(* PLC project HomeAutomation.ecp, WAGO e!COCKPIT e!COCKPIT *)
(* stored: creationDateTime 2023-02-09T18:04:59.3386506, modificationDateTime 2023-02-09T18:04:38.0443981 *)

{attribute 'to_string'}
TYPE Dimmer : (idle, soft_turn_on_restore, soft_turn_off, quick_turn_on, quick_turn_off, ramp_up_or_down, low_or_high_entering, low_or_high_leaving, low_or_high_released_by_user, blink);
END_TYPE

TYPE DIMMER_CURVE : (linear, logarithmic, cubic);
END_TYPE

TYPE MQTT_DISCOVERY_BASE : STRUCT
  name : JSONVAR;
  obj_id : JSONVAR;  (* object_id *)
  uniq_id : JSONVAR;  (* unique_id *)
  avty_t : JSONVAR;  (* availability_topic *)
  pl_avail : JSONVAR;  (* payload_available *)
  pl_not_avail : JSONVAR;  (* payload_not_available *)
  dev : MQTT_DISCOVERY_DEVICE;  (* device *)
  meta : JSONVAR;  (* extra metadata *)
END_STRUCT;
END_TYPE

TYPE MQTT_DISCOVERY_BINARY_SENSOR : STRUCT
  stat_t : JSONVAR;  (* state_topic *)
  pl_on : JSONVAR;  (* payload_on *)
  pl_off : JSONVAR;  (* payload_off *)
  dev_cla : JSONVAR;  (* device class *)
END_STRUCT;
END_TYPE

TYPE MQTT_DISCOVERY_COVER : STRUCT
  cmd_t : JSONVAR;  (* command_topic *)
  pl_open : JSONVAR;  (* payload open *)
  pl_cls : JSONVAR;  (* payload_close *)
  pl_stop : JSONVAR;  (* payload_stop *)
  stat_t : JSONVAR;  (* state topic *)
  stat_open : JSONVAR;  (* state open *)
  stat_clsd : JSONVAR;  (* state closed *)
  opt : JSONVAR;  (* optimistic *)
  dev_cla : JSONVAR;  (* device class *)
END_STRUCT;
END_TYPE

TYPE MQTT_DISCOVERY_DEVICE : STRUCT
  name : JSONVAR;
  cu : JSONVAR;  (* configuration_url *)
  ids : JSONVAR;  (* identifiers *)
  mf : JSONVAR;  (* manufacturer *)
  mdl : JSONVAR;  (* model *)
  sw : JSONVAR;  (* sw_version *)
  hw : JSONVAR;  (* hw_version *)
END_STRUCT;
END_TYPE

TYPE MQTT_DISCOVERY_LIGHT : STRUCT
  cmd_t : JSONVAR;  (* command_topic *)
  pl_on : JSONVAR;  (* payload_on *)
  pl_off : JSONVAR;  (* payload_off *)
  stat_t : JSONVAR;  (* state_topic *)
  opt : JSONVAR;  (* optimistic *)
END_STRUCT;
END_TYPE

TYPE MQTT_DISCOVERY_LIGHT_DIMMER : STRUCT
  bri_stat_t : JSONVAR;  (* brightness state topic *)
  bri_cmd_t : JSONVAR;  (* brightness command topic *)
  bri_scl : JSONVAR;  (* brightness scale *)
  on_cmd_type : JSONVAR;  (* on command type *)
  dmxChannel : JSONVAR;  (* DMX *)
  dmxWidth : JSONVAR;
  dmxUniverse : JSONVAR;
END_STRUCT;
END_TYPE

TYPE MQTT_DISCOVERY_LOCK : STRUCT
  cmd_t : JSONVAR;  (* command_topic *)
  pl_lock : JSONVAR;  (* payload lock *)
  pl_unlk : JSONVAR;  (* payload unlock *)
  stat_t : JSONVAR;  (* state_topic *)
  stat_locked : JSONVAR;  (* state locked *)
  stat_unlocked : JSONVAR;  (* state unlocked *)
  opt : JSONVAR;  (* optimistic *)
END_STRUCT;
END_TYPE

TYPE MQTT_DISCOVERY_SENSOR : STRUCT
  stat_t : JSONVAR;  (* state_topic *)
  exp_aft : JSONVAR;  (* expire after *)
END_STRUCT;
END_TYPE

TYPE MQTT_DISCOVERY_SIREN : STRUCT
  cmd_t : JSONVAR;  (* command_topic *)
  pl_on : JSONVAR;  (* payload_on *)
  pl_off : JSONVAR;  (* payload_off *)
  stat_t : JSONVAR;  (* state_topic *)
  stat_on : JSONVAR;  (* state on *)
  stat_off : JSONVAR;  (* state off *)
  opt : JSONVAR;  (* optimistic *)
END_STRUCT;
END_TYPE

TYPE MQTT_DISCOVERY_SWITCH : STRUCT
  cmd_t : JSONVAR;  (* command_topic *)
  pl_on : JSONVAR;  (* payload_on *)
  pl_off : JSONVAR;  (* payload_off *)
  stat_t : JSONVAR;  (* state_topic *)
  stat_on : JSONVAR;  (* state on *)
  stat_off : JSONVAR;  (* state off *)
  opt : JSONVAR;  (* optimistic *)
  dev_cla : JSONVAR;  (* device class *)
END_STRUCT;
END_TYPE

TYPE MQTT_MESSAGE : STRUCT
  Payload : STRING(1500);
  Topic : STRING(128);
  Qos : MQTT.QoS;
  MqttRetain : BOOL;
END_STRUCT;
END_TYPE

TYPE RS485_EASTRON_SDM_Devices : (SDM120, SDM220, SDM630);
END_TYPE

TYPE RS485_RtuQuery : STRUCT
  DeviceId : BYTE;
  FunctionCode : BYTE;
  ReadAddress : UINT;
  ReadQuantity : UINT;
  WriteAddress : UINT;
  WriteQuantity : UINT;
  WriteData : ARRAY[0..124] OF WORD;
END_STRUCT;
END_TYPE

TYPE VIRTUAL_MODES : (Input, Output);
END_TYPE

INTERFACE RS485Device
METHOD RequestBusTime : BOOL
END_METHOD
METHOD GetRtuQuery : RS485_RtuQuery
END_METHOD
METHOD ProcessDataArray
  VAR_INPUT
    Error : POINTER TO BOOL;
    Data : POINTER TO ARRAY[0..124] OF WORD;
  END_VAR
END_METHOD
END_INTERFACE

{attribute 'reflection'}
FUNCTION_BLOCK FB_BASE_MQTT_DISCOVERY_DEVICE
  VAR
    name : STRING;
    cu : STRING;  (* configuration_url *)
    cns : ARRAY[1..2] OF ARRAY[1..2] OF STRING;  (* connections *)
    ids : STRING;  (* identifiers *)
    mf : STRING;  (* manufacturer *)
    mdl : STRING;  (* model *)
    sw : STRING;  (* sw_version *)
    hw : STRING;  (* hw_version *)
    ip : STRING;
    mac : STRING;
    sAppName : STRING := 'Application';  (* must identic to the name in the device tree *)
    iecResult : RTS_IEC_RESULT;
    xInit : BOOL := TRUE;
    pApp : POINTER TO CmpApp.APPLICATION;
    stAppInfo : CmpApp.APPLICATION_INFO;
    pstAppInfo : POINTER TO CmpApp.APPLICATION_INFO := ADR(stAppInfo);
    {attribute 'instance-path'}
    {attribute 'noinit'}
    InstanceName : STRING;  (* object's full instance name *)
    Startup : BOOL := TRUE;
    InitMqttDone : BOOL;
    pMqttPublishQueue : POINTER TO FB_MqttPublishQueue;
    availabilityTopic : STRING;
    availabilityOnline : STRING;
    availabilityOffline : STRING;
    MqttDiscoveryPrefix : STRING;
    MqttDiscMsgBinSens : MQTT_DISCOVERY_BINARY_SENSOR;
    MqttDiscMsgCover : MQTT_DISCOVERY_COVER;
    MqttDiscMsgLightDim : MQTT_DISCOVERY_LIGHT_DIMMER;
    MqttDiscMsgLight : MQTT_DISCOVERY_LIGHT;
    MqttDiscMsgLock : MQTT_DISCOVERY_LOCK;
    MqttDiscMsgSensor : MQTT_DISCOVERY_SENSOR;
    MqttDiscMsgSiren : MQTT_DISCOVERY_SIREN;
    MqttDiscMsgSwitch : MQTT_DISCOVERY_SWITCH;
  END_VAR

            
          

{attribute 'reflection'}
METHOD CreateBinarySensorEntity
  VAR_INPUT
    Name : STRING;  (* default *)
    Id : STRING;
    Meta : STRING;
    StateTopic : STRING;  (* entity specific *)
    PayloadOn : STRING;
    PayloadOff : STRING;
    DeviceClass : STRING;
  END_VAR
  VAR
    EntityId : STRING(25) := 'binary_sensor';
    ComposeJSON : STRUCT_TO_JSON;
    MqttJSON : STRING(1500);
    MqttTopic : STRING(100);
  END_VAR
                  MqttTopic := CONCAT(CONCAT(CONCAT(CONCAT(THIS^.MqttDiscoveryPrefix, EntityId),'/'), Id),'/config' );


// 	Entity related: Basis
MqttDiscMsgBinSens.name.CharString :=  name; // friendly name
MqttDiscMsgBinSens.obj_id.CharString :=  Id; 
MqttDiscMsgBinSens.uniq_id.CharString :=  Id; 

// Entity related: Specific
MqttDiscMsgBinSens.stat_t.CharString := StateTopic;
MqttDiscMsgBinSens.pl_on.CharString := PayloadOn;
MqttDiscMsgBinSens.pl_off.CharString := PayloadOff;
MqttDiscMsgBinSens.dev_cla.CharString := DeviceClass;

// Availabilty related
MqttDiscMsgBinSens.avty_t.CharString :=  THIS^.availabilityTopic;
MqttDiscMsgBinSens.pl_avail.CharString :=   THIS^.availabilityOnline;
MqttDiscMsgBinSens.pl_not_avail.CharString :=  THIS^.availabilityOffline;

// Device related
MqttDiscMsgBinSens.dev.cu.CharString := THIS^.cu;
MqttDiscMsgBinSens.dev.name.CharString := THIS^.name;
MqttDiscMsgBinSens.dev.hw.CharString := THIS^.hw;
MqttDiscMsgBinSens.dev.ids.CharString := THIS^.ids;
MqttDiscMsgBinSens.dev.sw.CharString := THIS^.sw;
MqttDiscMsgBinSens.dev.mdl.CharString := THIS^.mdl;
MqttDiscMsgBinSens.dev.mf.CharString := THIS^.mf;
	
// Extra meta-data
IF NOT CommonTypesAndFunctions.StrEquals(str1:= ADR(meta), str2:= ADR('')) THEN
	MqttDiscMsgBinSens.meta.CharString := meta;
END_IF

ComposeJSON(
	JSONString:= ADR(MqttJSON), 
	JSONStringSize:= SIZEOF(MqttJSON),
	JSONVars:= ADR(MqttDiscMsgBinSens),
	NumberOfVars:= SIZEOF(MqttDiscMsgBinSens) / SIZEOF(JSONVAR),
	MaxLevel := 1,
);
ComposeJSON.Execute := TRUE;
ComposeJSON();

IF MqttJSON = '' THEN
	Mqttvariables.MQTT_logger.send(str:=CONCAT(CONCAT('ERROR ',Id), ' had empty MqttJSON'), instance := 'bla');
ELSIF NOT (MqttJSON = '') THEN
	pMqttPublishQueue^.AddMessage(
		Payload:= MqttJSON,
		Topic := MqttTopic,
		Qos := MQTT.QoS.ExactlyOnce,
		MqttRetain := TRUE,
	);
	Mqttvariables.MQTT_logger.send(str:=CONCAT(CONCAT('Added ',Id), ' as MQTT dicovery'), instance := 'bla');
END_IF

                
END_METHOD

METHOD CreateCoverEntity
  VAR_INPUT
    Name : STRING;  (* default *)
    Id : STRING;
    Meta : STRING;
    CommandTopic : STRING;  (* entity specific *)
    PayloadOpen : STRING;
    PayloadClose : STRING;
    PayloadStop : STRING;
    StateTopic : STRING;
    StateOpen : STRING;
    StateClosed : STRING;
    Deviceclass : STRING;
  END_VAR
  VAR
    EntityId : STRING(25) := 'cover';
    ComposeJSON : STRUCT_TO_JSON;
    MqttJSON : STRING(1500);
    MqttTopic : STRING(100);
  END_VAR
                  MqttTopic := CONCAT(CONCAT(CONCAT(CONCAT(THIS^.MqttDiscoveryPrefix, EntityId),'/'), Id),'/config' );

// 	Entity related: Basis
MqttDiscMsgCover.name.CharString :=  name; // friendly name
MqttDiscMsgCover.obj_id.CharString :=  Id; 
MqttDiscMsgCover.uniq_id.CharString :=  Id; 

// Entity related: Specific
MqttDiscMsgCover.cmd_t.CharString := CommandTopic;
MqttDiscMsgCover.pl_open.CharString := PayloadOpen;
MqttDiscMsgCover.pl_cls.CharString := PayloadClose;
MqttDiscMsgCover.pl_stop.CharString := PayloadStop;
MqttDiscMsgCover.stat_t.CharString := StateTopic;
MqttDiscMsgCover.stat_open.CharString := StateOpen;
MqttDiscMsgCover.stat_clsd.CharString := StateClosed;
MqttDiscMsgCover.opt.Boolean := FALSE;
MqttDiscMsgCover.dev_cla.CharString := Deviceclass;

// Availabilty related
MqttDiscMsgCover.avty_t.CharString :=  THIS^.availabilityTopic;
MqttDiscMsgCover.pl_avail.CharString :=   THIS^.availabilityOnline;
MqttDiscMsgCover.pl_not_avail.CharString :=  THIS^.availabilityOffline;

// Device related
MqttDiscMsgCover.dev.cu.CharString := THIS^.cu;
MqttDiscMsgCover.dev.name.CharString := THIS^.name;
MqttDiscMsgCover.dev.hw.CharString := THIS^.hw;
MqttDiscMsgCover.dev.ids.CharString := THIS^.ids;
MqttDiscMsgCover.dev.sw.CharString := THIS^.sw;
MqttDiscMsgCover.dev.mdl.CharString := THIS^.mdl;
MqttDiscMsgCover.dev.mf.CharString := THIS^.mf;
	
// Extra meta-data
IF NOT CommonTypesAndFunctions.StrEquals(str1:= ADR(meta), str2:= ADR('')) THEN
	MqttDiscMsgCover.meta.CharString := meta;
END_IF

ComposeJSON(
	JSONString:= ADR(MqttJSON), 
	JSONStringSize:= SIZEOF(MqttJSON),
	JSONVars:= ADR(MqttDiscMsgCover),
	NumberOfVars:= SIZEOF(MqttDiscMsgCover) / SIZEOF(JSONVAR),
	MaxLevel := 1,
);
ComposeJSON.Execute := TRUE;
ComposeJSON();

IF MqttJSON = '' THEN
	Mqttvariables.MQTT_logger.send(str:=CONCAT(CONCAT('ERROR ',Id), ' had empty MqttJSON'), instance := 'bla');
ELSIF NOT (MqttJSON = '') THEN
	pMqttPublishQueue^.AddMessage(
		Payload:= MqttJSON,
		Topic := MqttTopic,
		Qos := MQTT.QoS.ExactlyOnce,
		MqttRetain := TRUE,
	);
	Mqttvariables.MQTT_logger.send(str:=CONCAT(CONCAT('Added ',Id), ' as MQTT dicovery'), instance := 'bla');
END_IF

                
END_METHOD

METHOD initBaseDevice
  VAR_INPUT
    Name : STRING;
    ConfigurationUrl : STRING;
    Identifiers : STRING;
    Manufacturer : STRING;
    Model : STRING;
    SoftwareVersion : STRING;
    HardwareVersion : STRING;
    IpAddress : STRING := '';
    MacAddress : STRING := '';
    availabilityTopic : STRING;
    availabilityOnline : STRING;
    availabilityOffline : STRING;
    MqttDiscoveryPrefix : STRING;
    pMqttPublishQueue : POINTER TO FB_MqttPublishQueue;
  END_VAR
                  THIS^.availabilityTopic := availabilityTopic;
THIS^.availabilityOnline := availabilityOnline;
THIS^.availabilityOffline := availabilityOffline;
THIS^.pMqttPublishQueue := pMqttPublishQueue;
THIS^.MqttDiscoveryPrefix := MqttDiscoveryPrefix;

THIS^.name := Name;
THIS^.cu:= ConfigurationUrl;
THIS^.ids:= Identifiers;
THIS^.mf:= Manufacturer;
THIS^.mdl:= Model;
THIS^.hw:= HardwareVersion;
THIS^.ip := IpAddress;
THIS^.mac := MacAddress;




                
END_METHOD

METHOD CreateLightEntity
  VAR_INPUT
    Name : STRING;  (* default *)
    Id : STRING;
    Meta : STRING;
    CommandTopic : STRING;  (* entity specific *)
    PayloadOn : STRING;
    PayloadOff : STRING;
    StateTopic : STRING;
  END_VAR
  VAR
    EntityId : STRING(25) := 'light';
    ComposeJSON : STRUCT_TO_JSON;
    MqttJSON : STRING(1500);
    MqttTopic : STRING(100);
  END_VAR
                  MqttTopic := CONCAT(CONCAT(CONCAT(CONCAT(THIS^.MqttDiscoveryPrefix, EntityId),'/'), Id),'/config' );

// 	Entity related: Basis
MqttDiscMsgLight.name.CharString :=  name; // friendly name
MqttDiscMsgLight.obj_id.CharString :=  Id; 
MqttDiscMsgLight.uniq_id.CharString :=  Id; 

// Entity related: Specific
MqttDiscMsgLight.cmd_t.CharString := CommandTopic;
MqttDiscMsgLight.pl_on.CharString := PayloadOn;
MqttDiscMsgLight.pl_off.CharString := PayloadOff;
MqttDiscMsgLight.stat_t.CharString := StateTopic;
MqttDiscMsgLight.opt.Boolean := FALSE;

// Availabilty related
MqttDiscMsgLight.avty_t.CharString :=  THIS^.availabilityTopic;
MqttDiscMsgLight.pl_avail.CharString :=   THIS^.availabilityOnline;
MqttDiscMsgLight.pl_not_avail.CharString :=  THIS^.availabilityOffline;

// Device related
MqttDiscMsgLight.dev.cu.CharString := THIS^.cu;
MqttDiscMsgLight.dev.name.CharString := THIS^.name;
MqttDiscMsgLight.dev.hw.CharString := THIS^.hw;
MqttDiscMsgLight.dev.ids.CharString := THIS^.ids;
MqttDiscMsgLight.dev.sw.CharString := THIS^.sw;
MqttDiscMsgLight.dev.mdl.CharString := THIS^.mdl;
MqttDiscMsgLight.dev.mf.CharString := THIS^.mf;
	
// Extra meta-data
IF NOT CommonTypesAndFunctions.StrEquals(str1:= ADR(meta), str2:= ADR('')) THEN
	MqttDiscMsgLight.meta.CharString := meta;
END_IF

ComposeJSON(
	JSONString:= ADR(MqttJSON), 
	JSONStringSize:= SIZEOF(MqttJSON),
	JSONVars:= ADR(MqttDiscMsgLight),
	NumberOfVars:= SIZEOF(MqttDiscMsgLight) / SIZEOF(JSONVAR),
	MaxLevel := 1,
);
ComposeJSON.Execute := TRUE;
ComposeJSON();

IF MqttJSON = '' THEN
	Mqttvariables.MQTT_logger.send(str:=CONCAT(CONCAT('ERROR ',Id), ' had empty MqttJSON'), instance := 'bla');
ELSIF NOT (MqttJSON = '') THEN
	pMqttPublishQueue^.AddMessage(
		Payload:= MqttJSON,
		Topic := MqttTopic,
		Qos := MQTT.QoS.ExactlyOnce,
		MqttRetain := TRUE,
	);
	Mqttvariables.MQTT_logger.send(str:=CONCAT(CONCAT('Added ',Id), ' as MQTT dicovery'), instance := 'bla');
END_IF

                
END_METHOD

METHOD CreateLockEntity
  VAR_INPUT
    Name : STRING;  (* default *)
    Id : STRING;
    Meta : STRING;
    CommandTopic : STRING;  (* entity specific *)
    PayloadLock : STRING;
    PayloadUnlock : STRING;
    StateTopic : STRING;
    StateLocked : STRING;
    StateUnlocked : STRING;
  END_VAR
  VAR
    EntityId : STRING(25) := 'lock';
    ComposeJSON : STRUCT_TO_JSON;
    MqttJSON : STRING(1500);
    MqttTopic : STRING(100);
  END_VAR
                  MqttTopic := CONCAT(CONCAT(CONCAT(CONCAT(THIS^.MqttDiscoveryPrefix, EntityId),'/'), Id),'/config' );

// 	Entity related: Basis
MqttDiscMsgLock.name.CharString :=  name; // friendly name
MqttDiscMsgLock.obj_id.CharString :=  Id; 
MqttDiscMsgLock.uniq_id.CharString :=  Id; 

// Entity related: Specific
MqttDiscMsgLock.cmd_t.CharString := CommandTopic;
MqttDiscMsgLock.pl_lock.CharString := PayloadLock;
MqttDiscMsgLock.pl_unlk.CharString := PayloadUnlock;
MqttDiscMsgLock.stat_t.CharString := StateTopic;
MqttDiscMsgLock.stat_locked.CharString := StateLocked;
MqttDiscMsgLock.stat_unlocked.CharString := StateUnlocked;
MqttDiscMsgLock.opt.Boolean := FALSE;

// Availabilty related
MqttDiscMsgLock.avty_t.CharString :=  THIS^.availabilityTopic;
MqttDiscMsgLock.pl_avail.CharString :=   THIS^.availabilityOnline;
MqttDiscMsgLock.pl_not_avail.CharString :=  THIS^.availabilityOffline;

// Device related
MqttDiscMsgLock.dev.cu.CharString := THIS^.cu;
MqttDiscMsgLock.dev.name.CharString := THIS^.name;
MqttDiscMsgLock.dev.hw.CharString := THIS^.hw;
MqttDiscMsgLock.dev.ids.CharString := THIS^.ids;
MqttDiscMsgLock.dev.sw.CharString := THIS^.sw;
MqttDiscMsgLock.dev.mdl.CharString := THIS^.mdl;
MqttDiscMsgLock.dev.mf.CharString := THIS^.mf;
	
// Extra meta-data
IF NOT CommonTypesAndFunctions.StrEquals(str1:= ADR(meta), str2:= ADR('')) THEN
	MqttDiscMsgLock.meta.CharString := meta;
END_IF

ComposeJSON(
	JSONString:= ADR(MqttJSON), 
	JSONStringSize:= SIZEOF(MqttJSON),
	JSONVars:= ADR(MqttDiscMsgLock),
	NumberOfVars:= SIZEOF(MqttDiscMsgLock) / SIZEOF(JSONVAR),
	MaxLevel := 1,
);
ComposeJSON.Execute := TRUE;
ComposeJSON();

IF MqttJSON = '' THEN
	Mqttvariables.MQTT_logger.send(str:=CONCAT(CONCAT('ERROR ',Id), ' had empty MqttJSON'), instance := 'bla');
ELSIF NOT (MqttJSON = '') THEN
	pMqttPublishQueue^.AddMessage(
		Payload:= MqttJSON,
		Topic := MqttTopic,
		Qos := MQTT.QoS.ExactlyOnce,
		MqttRetain := TRUE,
	);
	Mqttvariables.MQTT_logger.send(str:=CONCAT(CONCAT('Added ',Id), ' as MQTT dicovery'), instance := 'bla');
END_IF

                
END_METHOD

METHOD CreateSirenEntity
  VAR_INPUT
    Name : STRING;  (* default *)
    Id : STRING;
    Meta : STRING;
    CommandTopic : STRING;  (* entity specific *)
    PayloadOn : STRING;
    PayloadOff : STRING;
    StateTopic : STRING;
    StateOnPayload : STRING;
    StateOffPayload : STRING;
  END_VAR
  VAR
    EntityId : STRING(25) := 'siren';
    ComposeJSON : STRUCT_TO_JSON;
    MqttJSON : STRING(1500);
    MqttTopic : STRING(100);
  END_VAR
                  MqttTopic := CONCAT(CONCAT(CONCAT(CONCAT(THIS^.MqttDiscoveryPrefix, EntityId),'/'), Id),'/config' );

// 	Entity related: Basis
MqttDiscMsgSiren.name.CharString :=  name; // friendly name
MqttDiscMsgSiren.obj_id.CharString :=  Id; 
MqttDiscMsgSiren.uniq_id.CharString :=  Id; 

// Entity related: Specific
MqttDiscMsgSiren.cmd_t.CharString := CommandTopic;
MqttDiscMsgSiren.pl_on.CharString := PayloadOn;
MqttDiscMsgSiren.pl_off.CharString := PayloadOff;
MqttDiscMsgSiren.stat_t.CharString := StateTopic;
MqttDiscMsgSiren.stat_on.CharString := StateOnPayload;
MqttDiscMsgSiren.stat_off.CharString := StateOffPayload;
MqttDiscMsgSiren.opt.Boolean := FALSE;

// Availabilty related
MqttDiscMsgSiren.avty_t.CharString :=  THIS^.availabilityTopic;
MqttDiscMsgSiren.pl_avail.CharString :=   THIS^.availabilityOnline;
MqttDiscMsgSiren.pl_not_avail.CharString :=  THIS^.availabilityOffline;

// Device related
MqttDiscMsgSiren.dev.cu.CharString := THIS^.cu;
MqttDiscMsgSiren.dev.name.CharString := THIS^.name;
MqttDiscMsgSiren.dev.hw.CharString := THIS^.hw;
MqttDiscMsgSiren.dev.ids.CharString := THIS^.ids;
MqttDiscMsgSiren.dev.sw.CharString := THIS^.sw;
MqttDiscMsgSiren.dev.mdl.CharString := THIS^.mdl;
MqttDiscMsgSiren.dev.mf.CharString := THIS^.mf;
	
// Extra meta-data
IF NOT CommonTypesAndFunctions.StrEquals(str1:= ADR(meta), str2:= ADR('')) THEN
	MqttDiscMsgSiren.meta.CharString := meta;
END_IF

ComposeJSON(
	JSONString:= ADR(MqttJSON), 
	JSONStringSize:= SIZEOF(MqttJSON),
	JSONVars:= ADR(MqttDiscMsgSiren),
	NumberOfVars:= SIZEOF(MqttDiscMsgSiren) / SIZEOF(JSONVAR),
	MaxLevel := 1,
);
ComposeJSON.Execute := TRUE;
ComposeJSON();

IF MqttJSON = '' THEN
	Mqttvariables.MQTT_logger.send(str:=CONCAT(CONCAT('ERROR ',Id), ' had empty MqttJSON'), instance := 'bla');
ELSIF NOT (MqttJSON = '') THEN
	pMqttPublishQueue^.AddMessage(
		Payload:= MqttJSON,
		Topic := MqttTopic,
		Qos := MQTT.QoS.ExactlyOnce,
		MqttRetain := TRUE,
	);
	Mqttvariables.MQTT_logger.send(str:=CONCAT(CONCAT('Added ',Id), ' as MQTT dicovery'), instance := 'bla');
END_IF

                
END_METHOD

METHOD CreateSensorEntity
  VAR_INPUT
    Name : STRING;  (* default *)
    Id : STRING;
    Meta : STRING;
    StateTopic : STRING;  (* entity specific *)
    ExpiryAfter : INT := 0;
  END_VAR
  VAR
    EntityId : STRING(25) := 'sensor';
    ComposeJSON : STRUCT_TO_JSON;
    MqttJSON : STRING(1500);
    MqttTopic : STRING(100);
  END_VAR
                  MqttTopic := CONCAT(CONCAT(CONCAT(CONCAT(THIS^.MqttDiscoveryPrefix, EntityId),'/'), Id),'/config' );

// 	Entity related: Basis
MqttDiscMsgSensor.name.CharString :=  name; // friendly name
MqttDiscMsgSensor.obj_id.CharString :=  Id; 
MqttDiscMsgSensor.uniq_id.CharString :=  Id; 

// Entity related: Specific
//MqttDiscoverySensorMessage.ic.CharString := Icon;
MqttDiscMsgSensor.stat_t.CharString := StateTopic;
MqttDiscMsgSensor.exp_aft.Integer := ExpiryAfter;

// Availabilty related
MqttDiscMsgSensor.avty_t.CharString :=  THIS^.availabilityTopic;
MqttDiscMsgSensor.pl_avail.CharString :=   THIS^.availabilityOnline;
MqttDiscMsgSensor.pl_not_avail.CharString :=  THIS^.availabilityOffline;

// Device related
MqttDiscMsgSensor.dev.cu.CharString := THIS^.cu;
MqttDiscMsgSensor.dev.name.CharString := THIS^.name;
MqttDiscMsgSensor.dev.hw.CharString := THIS^.hw;
MqttDiscMsgSensor.dev.ids.CharString := THIS^.ids;
MqttDiscMsgSensor.dev.sw.CharString := THIS^.sw;
MqttDiscMsgSensor.dev.mdl.CharString := THIS^.mdl;
MqttDiscMsgSensor.dev.mf.CharString := THIS^.mf;
	
// Extra meta-data
IF NOT CommonTypesAndFunctions.StrEquals(str1:= ADR(meta), str2:= ADR('')) THEN
	MqttDiscMsgSensor.meta.CharString := meta;
END_IF

ComposeJSON(
	JSONString:= ADR(MqttJSON), 
	JSONStringSize:= SIZEOF(MqttJSON),
	JSONVars:= ADR(MqttDiscMsgSensor),
	NumberOfVars:= SIZEOF(MqttDiscMsgSensor) / SIZEOF(JSONVAR),
	MaxLevel := 1,
);
ComposeJSON.Execute := TRUE;
ComposeJSON();

IF MqttJSON = '' THEN
	Mqttvariables.MQTT_logger.send(str:=CONCAT(CONCAT('ERROR ',Id), ' had empty MqttJSON'), instance := 'bla');
ELSIF NOT (MqttJSON = '') THEN
	pMqttPublishQueue^.AddMessage(
		Payload:= MqttJSON,
		Topic := MqttTopic,
		Qos := MQTT.QoS.ExactlyOnce,
		MqttRetain := TRUE,
	);
	Mqttvariables.MQTT_logger.send(str:=CONCAT(CONCAT('Added ',Id), ' as MQTT dicovery'), instance := 'bla');
END_IF

                
END_METHOD

METHOD CreateLightDimmerEntity
  VAR_INPUT
    Name : STRING;  (* default *)
    Id : STRING;
    Meta : STRING;
    CommandTopic : STRING;  (* entity specific *)
    PayloadOn : STRING;
    PayloadOff : STRING;
    StateTopic : STRING;
    BrightnessCommandTopic : STRING;
    BrightnessStateTopic : STRING;
    BrightnessScale : INT;
    DmxChannel : INT := 0;  (* dmx specific *)
    DmxWidth : INT := 0;
    DmxUniverse : INT := 0;
  END_VAR
  VAR
    EntityId : STRING(25) := 'light';
    ComposeJSON : STRUCT_TO_JSON;
    MqttJSON : STRING(1500);
    MqttTopic : STRING(100);
  END_VAR
                  MqttTopic := CONCAT(CONCAT(CONCAT(CONCAT(THIS^.MqttDiscoveryPrefix, EntityId),'/'), Id),'/config' );

// 	Entity related: Basis
MqttDiscMsgLightDim.name.CharString :=  name; // friendly name
MqttDiscMsgLightDim.obj_id.CharString :=  Id; 
MqttDiscMsgLightDim.uniq_id.CharString :=  Id; 

// Entity related: Specific
MqttDiscMsgLightDim.cmd_t.CharString := CommandTopic;
MqttDiscMsgLightDim.pl_on.CharString := PayloadOn;
MqttDiscMsgLightDim.pl_off.CharString := PayloadOff;
MqttDiscMsgLightDim.stat_t.CharString := StateTopic;
MqttDiscMsgLightDim.opt.Boolean := FALSE;

MqttDiscMsgLightDim.bri_cmd_t.CharString := BrightnessCommandTopic;
MqttDiscMsgLightDim.bri_stat_t.CharString := BrightnessStateTopic;
MqttDiscMsgLightDim.bri_scl.Integer := BrightnessScale;
MqttDiscMsgLightDim.on_cmd_type.CharString := 'last';

MqttDiscMsgLightDim.dmxChannel.Integer := DmxChannel;
MqttDiscMsgLightDim.dmxWidth.Integer := DmxWidth;
MqttDiscMsgLightDim.dmxUniverse.Integer := DmxUniverse;

// Availabilty related
MqttDiscMsgLightDim.avty_t.CharString :=  THIS^.availabilityTopic;
MqttDiscMsgLightDim.pl_avail.CharString :=   THIS^.availabilityOnline;
MqttDiscMsgLightDim.pl_not_avail.CharString :=  THIS^.availabilityOffline;

// Device related
MqttDiscMsgLightDim.dev.cu.CharString := THIS^.cu;
MqttDiscMsgLightDim.dev.name.CharString := THIS^.name;
MqttDiscMsgLightDim.dev.hw.CharString := THIS^.hw;
MqttDiscMsgLightDim.dev.ids.CharString := THIS^.ids;
MqttDiscMsgLightDim.dev.sw.CharString := THIS^.sw;
MqttDiscMsgLightDim.dev.mdl.CharString := THIS^.mdl;
MqttDiscMsgLightDim.dev.mf.CharString := THIS^.mf;
	
// Extra meta-data
IF NOT CommonTypesAndFunctions.StrEquals(str1:= ADR(meta), str2:= ADR('')) THEN
	MqttDiscMsgLightDim.meta.CharString := meta;
END_IF

ComposeJSON(
	JSONString:= ADR(MqttJSON), 
	JSONStringSize:= SIZEOF(MqttJSON),
	JSONVars:= ADR(MqttDiscMsgLightDim),
	NumberOfVars:= SIZEOF(MqttDiscMsgLightDim) / SIZEOF(JSONVAR),
	MaxLevel := 1,
);
ComposeJSON.Execute := TRUE;
ComposeJSON();

IF MqttJSON = '' THEN
	Mqttvariables.MQTT_logger.send(str:=CONCAT(CONCAT('ERROR ',Id), ' had empty MqttJSON'), instance := 'bla');
ELSIF NOT (MqttJSON = '') THEN
	pMqttPublishQueue^.AddMessage(
		Payload:= MqttJSON,
		Topic := MqttTopic,
		Qos := MQTT.QoS.ExactlyOnce,
		MqttRetain := TRUE,
	);
	Mqttvariables.MQTT_logger.send(str:=CONCAT(CONCAT('Added ',Id), ' as MQTT dicovery'), instance := 'bla');
END_IF

                
END_METHOD

METHOD CreateSwitchEntity
  VAR_INPUT
    Name : STRING;  (* default *)
    Id : STRING;
    Meta : STRING;
    CommandTopic : STRING;  (* entity specific *)
    PayloadOn : STRING;
    PayloadOff : STRING;
    StateTopic : STRING;
    StateOnPayload : STRING;
    StateOffPayload : STRING;
    DeviceClass : STRING;
  END_VAR
  VAR
    EntityId : STRING(25) := 'switch';
    ComposeJSON : STRUCT_TO_JSON;
    MqttJSON : STRING(1500);
    MqttTopic : STRING(100);
  END_VAR
                  MqttTopic := CONCAT(CONCAT(CONCAT(CONCAT(THIS^.MqttDiscoveryPrefix, EntityId),'/'), Id),'/config' );

// 	Entity related: Basis
MqttDiscMsgSwitch.name.CharString :=  name; // friendly name
MqttDiscMsgSwitch.obj_id.CharString :=  Id; 
MqttDiscMsgSwitch.uniq_id.CharString :=  Id; 

// Entity related: Specific
MqttDiscMsgSwitch.cmd_t.CharString := CommandTopic;
MqttDiscMsgSwitch.pl_on.CharString := PayloadOn;
MqttDiscMsgSwitch.pl_off.CharString := PayloadOff;
MqttDiscMsgSwitch.stat_t.CharString := StateTopic;
MqttDiscMsgSwitch.stat_on.CharString := StateOnPayload;
MqttDiscMsgSwitch.stat_off.CharString := StateOffPayload;
MqttDiscMsgSwitch.opt.Boolean := FALSE;
MqttDiscMsgSwitch.dev_cla.CharString := DeviceClass;

// Availabilty related
MqttDiscMsgSwitch.avty_t.CharString :=  THIS^.availabilityTopic;
MqttDiscMsgSwitch.pl_avail.CharString :=   THIS^.availabilityOnline;
MqttDiscMsgSwitch.pl_not_avail.CharString :=  THIS^.availabilityOffline;

// Device related
MqttDiscMsgSwitch.dev.cu.CharString := THIS^.cu;
MqttDiscMsgSwitch.dev.name.CharString := THIS^.name;
MqttDiscMsgSwitch.dev.hw.CharString := THIS^.hw;
MqttDiscMsgSwitch.dev.ids.CharString := THIS^.ids;
MqttDiscMsgSwitch.dev.sw.CharString := THIS^.sw;
MqttDiscMsgSwitch.dev.mdl.CharString := THIS^.mdl;
MqttDiscMsgSwitch.dev.mf.CharString := THIS^.mf;
	
// Extra meta-data
IF NOT CommonTypesAndFunctions.StrEquals(str1:= ADR(meta), str2:= ADR('')) THEN
	MqttDiscMsgSwitch.meta.CharString := meta;
END_IF

ComposeJSON(
	JSONString:= ADR(MqttJSON), 
	JSONStringSize:= SIZEOF(MqttJSON),
	JSONVars:= ADR(MqttDiscMsgSwitch),
	NumberOfVars:= SIZEOF(MqttDiscMsgSwitch) / SIZEOF(JSONVAR),
	MaxLevel := 1,
);
ComposeJSON.Execute := TRUE;
ComposeJSON();

IF MqttJSON = '' THEN
	Mqttvariables.MQTT_logger.send(str:=CONCAT(CONCAT('ERROR ',Id), ' had empty MqttJSON'), instance := 'bla');
ELSIF NOT (MqttJSON = '') THEN
	pMqttPublishQueue^.AddMessage(
		Payload:= MqttJSON,
		Topic := MqttTopic,
		Qos := MQTT.QoS.ExactlyOnce,
		MqttRetain := TRUE,
	);
	Mqttvariables.MQTT_logger.send(str:=CONCAT(CONCAT('Added ',Id), ' as MQTT dicovery'), instance := 'bla');
END_IF

                
END_METHOD
END_FUNCTION_BLOCK

{attribute 'reflection'}
FUNCTION_BLOCK FB_INPUT_BINARYSENSOR_MQTT EXTENDS FB_MQTT_BASE
  VAR_INPUT
    BS : BOOL;
  END_VAR
  VAR_OUTPUT
    Q : BOOL;  (* Follows the input but debounced *)
    EVENT : BOOL;  (* Event outputs only high for on clock cycle *)
    EVENT_R : BOOL;
    EVENT_F : BOOL;
  END_VAR
  VAR
    {attribute 'instance-path'}
    {attribute 'noinit'}
    InstancePath : STRING;  (* object's full instance name *)
    Startup : BOOL := TRUE;
    FB_DEBOUNCE : OSCAT_BUILDING.DEBOUNCE;  (* to debounce the physical input *)
    FB_R_TRIG : Standard.R_TRIG;  (* to detect a rising edge on the debounced signal *)
    FB_F_TRIG : Standard.F_TRIG;  (* to detect a falling edge on the debounced signal *)
    T_TurnOffDelay : TIME := TIME#0ms;
    FB_TurnOffDelayTimer : TOF;
    MqttDiscoveryMessage : MQTT_DISCOVERY_BINARY_SENSOR;
  END_VAR

            FB_DEBOUNCE(IN := BS,	
	TD := T#50MS, (* 2x cyle + 10ms *)
	PM := FALSE
	);
	
FB_TurnOffDelayTimer(IN:=FB_DEBOUNCE.Q,
	PT := T_TurnOffDelay,
	Q=>Q
	);

FB_R_TRIG(CLK := FB_TurnOffDelayTimer.Q);
FB_F_TRIG(CLK := FB_TurnOffDelayTimer.Q);

EVENT := FB_R_TRIG.Q OR FB_F_TRIG.Q;
EVENT_R := FB_R_TRIG.Q;
EVENT_F := FB_F_TRIG.Q;

IF (FB_R_TRIG.Q OR (Startup AND FB_DEBOUNCE.Q)) AND InitMqttDone THEN
	pMqttPublishQueue^.AddMessage(
		Payload := 'ON',
		Topic := CONCAT(MqttPublishTopicPrefix^, MqttPublishTopicSuffix),
		Qos := MQTT.QoS.ExactlyOnce,
		MqttRetain := TRUE
	);
	Startup:=FALSE;	
END_IF

IF (FB_F_TRIG.Q OR (Startup AND NOT(FB_DEBOUNCE.Q))) AND InitMqttDone THEN
	pMqttPublishQueue^.AddMessage(
		Payload := 'OFF',
		Topic := CONCAT(MqttPublishTopicPrefix^, MqttPublishTopicSuffix),
		Qos := MQTT.QoS.ExactlyOnce,
		MqttRetain := TRUE
	);
	Startup:=FALSE;	
END_IF
          

METHOD InitMqtt
  VAR_INPUT
    MQTTPublishPrefix : POINTER TO STRING;
    pMqttPublishQueue : POINTER TO FB_MqttPublishQueue;
  END_VAR
                  SUPER^._InstancePath := THIS^.InstancePath; // Due to reflection its location is important

(*pass trough*)
THIS^.pMqttPublishQueue := pMqttPublishQueue;
THIS^.MqttPublishTopicPrefix:=MQTTPublishPrefix;
SUPER^.InitBaseMqtt();

                
END_METHOD

METHOD InitMqttDiscovery
  VAR_INPUT
    Device : POINTER TO FB_PLC_MQTT_DISCOVERY_DEVICE;
    Name : STRING(255);
    DeviceClass : STRING(100) := 'smoke';
    overruleId : STRING(255) := '';
    meta : STRING(255) := '';
  END_VAR
  VAR
    id : STRING(255);
  END_VAR
                  IF InitMqttDone AND NOT initMqttDiscoveryDone THEN
	
	IF CommonTypesAndFunctions.StrEquals(str1:= ADR(overruleId), str2:= ADR('')) THEN
		id := CONCAT(CONCAT(THIS^.DeviceName,'_'), THIS^.InstanceNamePt^); // 'FB_DI_PB_003'
	ELSE
		id := overruleId; // 'MY_PH_GND_HALL_01'
	END_IF
	
	Device^.CreateBinarySensorEntity(
		Id := id,
		Name := name,
		Meta := meta,
		StateTopic := THIS^.MQTTPublishTopic,
		PayloadOn := 'ON',
		PayloadOff := 'OFF',
		DeviceClass := DeviceClass);
		
	initMqttDiscoveryDone := TRUE;
END_IF		
                
END_METHOD

METHOD ConfigureFunctionBlock
  VAR_INPUT
    T_TurnOffDelay : TIME;
  END_VAR
                  THIS^.T_TurnOffDelay:=T_TurnOffDelay;
                
END_METHOD
END_FUNCTION_BLOCK

{attribute 'reflection'}
FUNCTION_BLOCK FB_INPUT_PUSHBUTTON_DIMMER_MQTT
  VAR_INPUT
    PB : BOOL;
    SET : BOOL;
    VAL : BYTE;
    RST : BOOL;
  END_VAR
  VAR_OUTPUT
    DIM : BYTE;
    DBL : BOOL;
    Q : BOOL;
    SINGLE : BOOL;
    DOUBLE : BOOL;
    LONG : BOOL;
    P_LONG : BOOL;
  END_VAR
  VAR
    {attribute 'instance-path'}
    {attribute 'noinit'}
    InstanceName : STRING;  (* object's full instance name *)
    InitMqttDone : BOOL;
    MqttPublishTopicPrefix : POINTER TO STRING;
    MqttPublishTopicSuffix : STRING(50);
    pMqttPublishQueue : POINTER TO FB_MqttPublishQueue;
    FB_DIMMER : OSCAT_BUILDING.DIMM_I;
    OutputDimmer : BOOL;
    Qos_Dimm : MQTT.QoS;
    Delta_Dimm : INT;
    FB_DETECTPUSH : OSCAT_BUILDING.CLICK_MODE;
    P_LONG_R_TRIG : Standard.R_TRIG;
    P_LONG_F_TRIG : Standard.F_TRIG;
    PreviousDim : BYTE;  (* Vars to detect statechanges on outputs *)
    PreviousQ : BOOL;
    PreviousDBL : BOOL;
    T_Debounce : TIME := TIME#10ms;  (* Default values for dimmer, can be overwritten by method call *)
    T_Reconfig : TIME := TIME#10s0ms;
    T_On_Max : TIME := TIME#0ms;
    T_Dimm_Start : TIME := TIME#400ms;
    T_Dimm : TIME := TIME#3s0ms;
    Min_On : BYTE := 50;
    Max_On : BYTE := 255;
    Soft_Dimm : BOOL := TRUE;
    Dbl_Toggle : BOOL := FALSE;
    Rst_Out : BOOL := FALSE;
    T_Long : TIME := TIME#400ms;  (* Default value for click mode, can be overwritten by method call *)
  END_VAR

            FB_DIMMER(
	IN:= PB,
	SET:= SET,
	VAL:= VAL,
	RST:= RST,
	OUT:= DIM,
	T_DEBOUNCE:= T_Debounce,
	T_RECONFIG:= T_Reconfig,
	T_ON_MAX:= T_On_Max,
	T_DIMM_START:= T_Dimm_Start,
	T_DIMM:= T_Dimm,
	MIN_ON:= Min_On,
	MAX_ON:= Max_On,
	SOFT_DIMM:= Soft_Dimm,
	DBL_TOGGLE:= Dbl_Toggle,
	RST_OUT:= Rst_Out,
	Q=> Q,
	DBL=> DBL);
	
FB_DETECTPUSH(
	IN:= PB, 	
	SINGLE=> SINGLE, 
	DOUBLE=> DOUBLE, 
	TP_LONG=> LONG, 
	T_LONG:= T_long);
	
P_LONG_R_TRIG(CLK:=FB_DETECTPUSH.LONG);
P_LONG_F_TRIG(CLK:=FB_DETECTPUSH.LONG);
	
IF (ABS(BYTE_TO_INT(PreviousDim) - BYTE_TO_INT(DIM)) >= Delta_Dimm OR PB = FALSE) AND DIM <> PreviousDim AND OutputDimmer AND InitMqttDone  THEN
	PreviousDim:=DIM;
	pMqttPublishQueue^.AddMessage(		
		Payload := BYTE_TO_STRING(DIM),
		Topic := CONCAT(CONCAT(MqttPublishTopicPrefix^, MqttPublishTopicSuffix), '/DIM'),
		Qos := MQTT.QoS.ExactlyOnce,
		MqttRetain := FALSE
	);
END_IF

IF FB_DIMMER.Q <> PreviousQ AND InitMqttDone THEN
	PreviousQ:=FB_DIMMER.Q;
	pMqttPublishQueue^.AddMessage(
		Payload := BOOL_TO_STRING(FB_DIMMER.Q),
		Topic := CONCAT(CONCAT(MqttPublishTopicPrefix^, MqttPublishTopicSuffix), '/Q'),
		Qos := Qos_Dimm,
		MqttRetain := TRUE
	);
END_IF

IF FB_DIMMER.DBL <> PreviousDBL AND InitMqttDone THEN
	PreviousDBL:=FB_DIMMER.DBL;
	pMqttPublishQueue^.AddMessage(
		Payload := BOOL_TO_STRING(FB_DIMMER.DBL),
		Topic := CONCAT(CONCAT(MqttPublishTopicPrefix^, MqttPublishTopicSuffix), '/DBL'),
		Qos := MQTT.QoS.ExactlyOnce,
		MqttRetain := TRUE
	);
END_IF

IF FB_DETECTPUSH.SINGLE AND InitMqttDone THEN
	pMqttPublishQueue^.AddMessage(
		Payload := 'SINGLE',
		Topic := CONCAT(MqttPublishTopicPrefix^, MqttPublishTopicSuffix),
		Qos := MQTT.QoS.ExactlyOnce,
		MqttRetain := FALSE
	);
END_IF

IF FB_DETECTPUSH.DOUBLE AND InitMqttDone THEN
	pMqttPublishQueue^.AddMessage(
		Payload := 'DOUBLE',
		Topic := CONCAT(MqttPublishTopicPrefix^, MqttPublishTopicSuffix),
		Qos := MQTT.QoS.ExactlyOnce,
		MqttRetain := FALSE
	);
END_IF

IF FB_DETECTPUSH.TP_LONG AND InitMqttDone THEN
	pMqttPublishQueue^.AddMessage(
		Payload := 'LONG',
		Topic := CONCAT(MqttPublishTopicPrefix^, MqttPublishTopicSuffix),
		Qos := MQTT.QoS.ExactlyOnce,
		MqttRetain := FALSE
	);
END_IF

IF (P_LONG_R_TRIG.Q OR P_LONG_F_TRIG.Q) AND InitMqttDone THEN
	pMqttPublishQueue^.AddMessage(
		Payload := BOOL_TO_STRING(FB_DETECTPUSH.LONG),
		Topic := CONCAT(CONCAT(MqttPublishTopicPrefix^, MqttPublishTopicSuffix),'/P_LONG'),
		Qos := MQTT.QoS.ExactlyOnce,
		MqttRetain := TRUE
	);
END_IF
          

METHOD InitMqtt
  VAR_INPUT
    MQTTPublishPrefix : POINTER TO STRING;
    pMqttPublishQueue : POINTER TO FB_MqttPublishQueue;
    OutputDimmer : BOOL;
    Qos_Dimm : MQTT.QoS;
    Delta_Dimm : INT;
  END_VAR
  VAR
    InstanceNamePt : POINTER TO STRING;
  END_VAR
                  THIS^.pMqttPublishQueue := pMqttPublishQueue;
THIS^.MqttPublishTopicPrefix := MQTTPublishPrefix;

InstanceNamePt := CommonTypesAndFunctions.FindLastDot(ADR(THIS^.InstanceName)) + 1;
THIS^.MqttPublishTopicSuffix := InstanceNamePt^;

THIS^.OutputDimmer:=OutputDimmer;
THIS^.Qos_Dimm:=Qos_Dimm;
THIS^.Delta_Dimm:=Delta_Dimm;

InitMqttDone := TRUE;
                
END_METHOD

METHOD ConfigureFunctionBlock
  VAR_INPUT
    T_Debounce : TIME;  (* Default values for dimmer, can be overwritten by method call *)
    T_Reconfig : TIME;
    T_On_Max : TIME;
    T_Dimm_Start : TIME;
    T_Dimm : TIME;
    Min_On : BYTE;
    Max_On : BYTE;
    Soft_Dimm : BOOL;
    Dbl_Toggle : BOOL;
    Rst_Out : BOOL;
    T_Long : TIME;  (* Default value for click mode, can be overwritten by method call *)
  END_VAR
                  THIS^.T_Debounce:=T_Debounce;
THIS^.T_Reconfig:=T_Reconfig;
THIS^.T_On_Max:=T_On_Max;
THIS^.T_Dimm_Start:=T_Dimm_Start;
THIS^.T_Dimm:=T_Dimm;
THIS^.Min_On:=Min_On;
THIS^.Max_On:=Max_On;

THIS^.T_Long:=T_Long;
                
END_METHOD
END_FUNCTION_BLOCK

{attribute 'reflection'}
FUNCTION_BLOCK FB_INPUT_PUSHBUTTON_MQTT EXTENDS FB_MQTT_BASE
  VAR_INPUT
    PB : BOOL;
  END_VAR
  VAR_OUTPUT
    SINGLE : BOOL;
    DOUBLE : BOOL;
    LONG : BOOL;
    P_LONG : BOOL;
  END_VAR
  VAR
    {attribute 'instance-path'}
    {attribute 'noinit'}
    InstancePath : STRING;  (* Refelection: object's full instance name *)
    FB_DETECTPUSH : OSCAT_BUILDING.CLICK_MODE;
    P_LONG_R_TRIG : Standard.R_TRIG;
    P_LONG_F_TRIG : Standard.F_TRIG;
    T_Long : TIME := TIME#400ms;  (* Default value for click mode, can be overwritten by method call *)
    MqttDiscoveryMessage : MQTT_DISCOVERY_SENSOR;
  END_VAR

            FB_DETECTPUSH(
	IN:= PB, 	
	SINGLE=> SINGLE, 
	DOUBLE=> DOUBLE, 
	TP_LONG=> LONG, 
	LONG=> P_LONG,
	T_LONG:= T_Long);
	
P_LONG_R_TRIG(CLK:=FB_DETECTPUSH.LONG);
P_LONG_F_TRIG(CLK:=FB_DETECTPUSH.LONG);
	
IF FB_DETECTPUSH.SINGLE AND InitMqttDone THEN
	pMqttPublishQueue^.AddMessage(
		Payload := 'SINGLE',
		Topic := CONCAT(MqttPublishTopicPrefix^, MqttPublishTopicSuffix),
		Qos := MQTT.QoS.ExactlyOnce,
		MqttRetain := FALSE
	);
END_IF

IF FB_DETECTPUSH.DOUBLE AND InitMqttDone THEN
	pMqttPublishQueue^.AddMessage(
		Payload := 'DOUBLE',
		Topic := CONCAT(MqttPublishTopicPrefix^, MqttPublishTopicSuffix),
		Qos := MQTT.QoS.ExactlyOnce,
		MqttRetain := FALSE
	);
END_IF

IF FB_DETECTPUSH.TP_LONG AND InitMqttDone THEN
	pMqttPublishQueue^.AddMessage(
		Payload := 'LONG',
		Topic := MQTTPublishTopic,
		Qos := MQTT.QoS.ExactlyOnce,
		MqttRetain := FALSE
	);
END_IF

IF P_LONG_F_TRIG.Q AND InitMqttDone THEN
	pMqttPublishQueue^.AddMessage(
		Payload := 'RELEASED',
		Topic := MQTTPublishTopic,
		Qos := MQTT.QoS.ExactlyOnce,
		MqttRetain := FALSE
	);
END_IF



IF (P_LONG_R_TRIG.Q OR P_LONG_F_TRIG.Q) AND InitMqttDone THEN
	

	pMqttPublishQueue^.AddMessage(
		Payload := BOOL_TO_STRING(FB_DETECTPUSH.LONG),
		Topic := CONCAT(MQTTPublishTopic,'/P_LONG'),
		Qos := MQTT.QoS.ExactlyOnce,
		MqttRetain := TRUE
	);
END_IF
          

METHOD InitMqttDiscovery
  VAR_INPUT
    Device : POINTER TO FB_PLC_MQTT_DISCOVERY_DEVICE;
    Name : STRING(255);
    overruleId : STRING(255) := '';
    meta : STRING(255) := '';
  END_VAR
  VAR
    id : STRING(255);
  END_VAR
                  IF InitMqttDone AND NOT initMqttDiscoveryDone THEN
	
	IF CommonTypesAndFunctions.StrEquals(str1:= ADR(overruleId), str2:= ADR('')) THEN
		id := CONCAT(CONCAT(THIS^.DeviceName,'_'), THIS^.InstanceNamePt^); // 'FB_DI_PB_003'
	ELSE
		id := overruleId; // 'MY_PH_GND_HALL_01'
	END_IF
	
	Device^.CreateSensorEntity(
		Name := name,
		Id := id,
		Meta := meta,
		StateTopic := THIS^.MQTTPublishTopic,
		ExpiryAfter := 2);

	initMqttDiscoveryDone := TRUE;
END_IF		
                
END_METHOD

METHOD InitMqtt
  VAR_INPUT
    MQTTPublishPrefix : POINTER TO STRING;
    pMqttPublishQueue : POINTER TO FB_MqttPublishQueue;
  END_VAR
                  SUPER^._InstancePath := THIS^.InstancePath; // Due to reflection its location is important

(*pass trough*)
THIS^.pMqttPublishQueue := pMqttPublishQueue;
THIS^.MqttPublishTopicPrefix:=MQTTPublishPrefix;
SUPER^.InitBaseMqtt();

                
END_METHOD

METHOD ConfigureFunctionBlock
  VAR_INPUT
    T_Long : TIME;  (* Default value for click mode, can be overwritten by method call *)
  END_VAR
                  THIS^.T_Long:=T_Long;
                
END_METHOD
END_FUNCTION_BLOCK

FUNCTION_BLOCK FB_MQTT_BASE
  VAR
    _InstancePath : STRING;
    InstanceNamePt : POINTER TO STRING;
    DeviceName : STRING;
    InitMqttDone : BOOL;
    MqttPublishTopicPrefix : POINTER TO STRING;  (* Publish (Out); *)
    MqttPublishTopicSuffix : STRING(50);
    MQTTPublishTopic : STRING(100);
    MqttSubscribeTopicPrefix : POINTER TO STRING;  (* Subscribe (In) *)
    MqttSubscribeTopicSuffix : STRING(50);
    MQTTSubscribeTopic : STRING(100);
    pMqttPublishQueue : POINTER TO FB_MqttPublishQueue;
    MqttHighRequest : BOOL;
    MqttLowRequest : BOOL;
    MqttQos : MQTT.QoS := MQTT.QoS.ExactlyOnce;
    MqttRetain : BOOL := TRUE;
    ComposeJSON : STRUCT_TO_JSON;  (* HA Discovery specific *)
    initMqttDiscoveryDone : BOOL := FALSE;
  END_VAR

            
          

METHOD InitBaseMqtt
  VAR
    MQTTPublishPrefix : POINTER TO STRING;
    MQTTSubscribePrefix : POINTER TO STRING;
    pMqttPublishQueue : POINTER TO FB_MqttPublishQueue;
  END_VAR
                  
(*Define instance names*)
InstanceNamePt := CommonTypesAndFunctions.FindLastDot(ADR(_InstancePath)) + 1;

DeviceName := LEFT(_InstancePath,find(_InstancePath, '.' )-1  ) ;

// Publish (Out);
IF	NOT CommonTypesAndFunctions.StrEquals(ADR(MqttPublishTopicPrefix),ADR('')) THEN
	THIS^.MqttPublishTopicSuffix := InstanceNamePt^;
	THIS^.MQTTPublishTopic := CONCAT(MqttPublishTopicPrefix^, THIS^.MqttPublishTopicSuffix);
END_IF

// Subscribe (In)
IF	NOT CommonTypesAndFunctions.StrEquals(ADR(MqttSubscribeTopicPrefix),ADR('')) THEN
	THIS^.MQTTSubscribeTopicSuffix := InstanceNamePt^;
	THIS^.MQTTSubscribeTopic := CONCAT(MqttSubscribeTopicPrefix^ ,THIS^.MQTTSubscribeTopicSuffix);
END_IF

InitMqttDone := TRUE;
                
END_METHOD
END_FUNCTION_BLOCK

FUNCTION_BLOCK FB_MQTT_LOG EXTENDS FB_MQTT_BASE
  VAR
    InstancePath : STRING := '.plc_log';  (* should have a dot in the name *)
    MqttDiscoveryMessage : MQTT_DISCOVERY_SENSOR;
  END_VAR

            
          

METHOD InitMqttDiscovery
  VAR_INPUT
    Device : POINTER TO FB_PLC_MQTT_DISCOVERY_DEVICE;
    Name : STRING(255) := 'plc_log';
    overruleId : STRING(255) := '';
    meta : STRING(255) := '';
  END_VAR
  VAR
    id : STRING(255);
  END_VAR
                  IF InitMqttDone AND NOT initMqttDiscoveryDone THEN
	
	IF CommonTypesAndFunctions.StrEquals(str1:= ADR(overruleId), str2:= ADR('')) THEN
		id := CONCAT(CONCAT(THIS^.DeviceName,'_'), THIS^.InstanceNamePt^); // 'FB_DI_PB_003'
	ELSE
		id := overruleId; // 'MY_PH_GND_HALL_01'
	END_IF	
	
	Device^.CreateSensorEntity(
		Name := name,
		Id := id,
		Meta := meta,
		StateTopic := THIS^.MQTTPublishTopic);

	initMqttDiscoveryDone := TRUE;
END_IF		
                
END_METHOD

METHOD send
  VAR_INPUT
    str : STRING(128);
    instance : STRING := '';
  END_VAR
                  IF InitMqttDone THEN
	pMqttPublishQueue^.AddMessage(
		Payload:= CONCAT(CONCAT(instance,' | '),str),
		Topic := THIS^.MQTTPublishTopic,
		Qos := 1,
		MqttRetain := TRUE
	);
END_IF		
                
END_METHOD

METHOD InitMqtt
  VAR_INPUT
    MQTTPublishPrefix : POINTER TO STRING;
    pMqttPublishQueue : POINTER TO FB_MqttPublishQueue;
    MqttQos : MQTT.QoS := MQTT.QoS.ExactlyOnce;
    MqttRetain : BOOL := FALSE;
  END_VAR
                  SUPER^._InstancePath := THIS^.InstancePath; // Due to reflection its location is important

(*pass trough*)
THIS^.pMqttPublishQueue := pMqttPublishQueue;
THIS^.MqttPublishTopicPrefix:=MQTTPublishPrefix;
THIS^.pMqttPublishQueue:=pMqttPublishQueue;

THIS^.MqttQos := MqttQos;
THIS^.MqttRetain := MqttRetain;

SUPER^.InitBaseMqtt();
                
END_METHOD
END_FUNCTION_BLOCK

FUNCTION_BLOCK FB_MqttPublishQueue
  VAR_OUTPUT
    EMPTY : BOOL := TRUE;
    FULL : BOOL;
  END_VAR
  VAR
    localMessage : MQTT_MESSAGE;
    fifo : ARRAY[0..n] OF MQTT_MESSAGE;
    pr : INT;
    pw : INT;
  END_VAR
  VAR CONSTANT
    n : INT := 1024;  (* changing this value will chage the number of stored elements in the fifo *)
  END_VAR

            
          

METHOD GetMessage : MQTT_MESSAGE
                  IF NOT EMPTY THEN
	GetMessage := fifo[pr];
	pr := OSCAT_BASIC.INC1(pr,n);
	EMPTY := pr = pw;
	FULL := FALSE;
END_IF;
                
END_METHOD

METHOD AddMessage
  VAR_INPUT
    Payload : STRING(1500);
    Topic : STRING(128);
    Qos : MQTT.QoS;
    MqttRetain : BOOL;
  END_VAR
                  IF NOT FULL THEN
	localMessage.Payload := Payload;
	localMessage.Topic := Topic;
	localMessage.Qos := Qos;
	localMessage.MqttRetain := MqttRetain;
	fifo[pw] := localMessage;
	pw := OSCAT_BASIC.INC1(pw,n);
	FULL := pw = pr;
	EMPTY := FALSE;
END_IF;
                
END_METHOD

METHOD Reset
                  pw := pr;
FULL := FALSE;
EMPTY := TRUE;
                
END_METHOD
END_FUNCTION_BLOCK

FUNCTION_BLOCK FB_MqttPublishWorker
  VAR_OUTPUT
    SendDone : BOOL;
  END_VAR
  VAR
    LocalMqttMessage : MQTT_MESSAGE;
    InitDone : BOOL;
    RequestToSend : BOOL;
    Send : BOOL;
    publish : MQTT.MQTTPublish;
  END_VAR

            //need to call publish here because of FB nums
publish(
	Topic:= ADR(LocalMqttMessage.Topic), 
	PayloadString:= ADR(LocalMqttMessage.Payload), 
	PublishAsString:= TRUE, 
	QoSIn:= LocalMqttMessage.Qos, 
	MRetain:= LocalMqttMessage.MqttRetain, 
	send:= Send);
	
IF NOT InitDone THEN RETURN; END_IF

IF RequestToSend THEN
	Send := TRUE;
	SendDone := FALSE;
END_IF

IF publish.done THEN
	 SendDone := TRUE;
	 RequestToSend:=FALSE;
	 Send:=FALSE;
END_IF
          

METHOD Init
  VAR_INPUT
    inputMQTT_IN_OUT : POINTER TO MQTT.MQTT_IN_OUT;  (* Pointer MQTTT exchange strucure *)
  END_VAR
                  publish.SetMqttInOut(MQTT_IN_OUT := inputMQTT_IN_OUT^);

InitDone := TRUE;
SendDone := TRUE;

                
END_METHOD

METHOD PublishMessage
  VAR_INPUT
    MqttMessage : MQTT_MESSAGE;
  END_VAR
                  LocalMqttMessage := MqttMessage;

RequestToSend:=TRUE;
                
END_METHOD
END_FUNCTION_BLOCK

{attribute 'reflection'}
FUNCTION_BLOCK FB_OUTPUT_BINARY_MQTT EXTENDS FB_MQTT_BASE IMPLEMENTS MQTT.MQTT_SUBSCRIBE_CALLBACK
  VAR_INPUT
    PRIO_HIGH : BOOL := FALSE;
    PRIO_LOW : BOOL := FALSE;
    TOGGLE : BOOL := FALSE;
  END_VAR
  VAR_OUTPUT
    OUT : BOOL;
  END_VAR
  VAR
    {attribute 'instance-path'}
    {attribute 'noinit'}
    InstancePath : STRING;  (* Refelection: object's full instance name *)
    Startup : BOOL := TRUE;
    MqttDiscMsgSwitch : MQTT_DISCOVERY_SWITCH;  (* ComposeJSONLight : STRUCT_TO_JSON; MqttDiscoveryMessageLight: MQTT_DISCOVERY_LIGHT; ComposeJSONLock : STRUCT_TO_JSON; MqttDiscoveryMessageLock: MQTT_DISCOVERY_LOCK; ComposeJSONSiren : STRUCT_TO_JSON; MqttDiscoveryMessageSiren: MQTT_DISCOVERY_SIREN; ComposeJSONSwitch : STRUCT_TO_JSON; *)
  END_VAR
  VAR PERSISTENT
    PreviousState : BOOL;  (* To retain output state through powercycles *)
  END_VAR

            IF Startup THEN
	OUT := PreviousState;
END_IF

IF PRIO_HIGH THEN
	OUT:=TRUE;
ELSIF(PRIO_LOW AND NOT (PRIO_HIGH)) THEN
	OUT:= FALSE;
ELSIF MqttHighRequest THEN
	OUT:= TRUE;
	MqttHighRequest := FALSE;
	MqttLowRequest := FALSE;
ELSIF MqttLowRequest THEN
	OUT:= FALSE;
	MqttHighRequest := FALSE;
	MqttLowRequest := FALSE;
ELSIF(TOGGLE) THEN
	OUT:=NOT(OUT);
END_IF;

IF ((PreviousState <> OUT) OR Startup) AND InitMqttDone THEN
	pMqttPublishQueue^.AddMessage(
		Payload := BOOL_TO_STRING(OUT),
		Topic := MQTTPublishTopic,
		Qos := MQTT.QoS.ExactlyOnce,
		MqttRetain := TRUE
	);	
	Startup:=FALSE;
END_IF	

PreviousState := OUT;
          

METHOD InitMqtt
  VAR_INPUT
    MQTTPublishPrefix : POINTER TO STRING;
    MQTTSubscribePrefix : POINTER TO STRING;
    pMqttPublishQueue : POINTER TO FB_MqttPublishQueue;
    pMqttCallbackCollector : POINTER TO MQTT.CallbackCollector;
  END_VAR
                  SUPER^._InstancePath := THIS^.InstancePath; // Due to reflection its location is important

(*pass trough*)
THIS^.pMqttPublishQueue := pMqttPublishQueue;
THIS^.MqttPublishTopicPrefix:=MQTTPublishPrefix;
THIS^.MQTTSubscribeTopicPrefix:=MQTTSubscribePrefix;
THIS^.pMqttPublishQueue:=pMqttPublishQueue;

SUPER^.InitBaseMqtt();
pMqttCallbackCollector^.put(instance:= THIS^); // register the FB agains the collector so mqtt events can be received


                
END_METHOD

METHOD PublishReceived : BOOL
  VAR_INPUT
    Data : MQTT.CALLBACK_DATA;  (* Collection of recived Data *)
  END_VAR
                  //first check if Mqtt is initialized, otherwise do nothing
IF NOT(InitMqttDone) THEN
	//mark the interface call from the collector as done
	PublishReceived := TRUE;
//check if the packet is for this FB
ELSIF CommonTypesAndFunctions.StrEquals(str1:= ADR(MQTTSubscribeTopic), str2:= Data.TopicOut) THEN
	//mark the interface call from the collector as done
	PublishReceived := TRUE;
	//now process the data
	IF FIND(Data.PayloadString^, 'TRUE') > 0 THEN
		MqttHighRequest := TRUE;
	END_IF
	IF FIND(Data.PayloadString^, 'FALSE') > 0 THEN
		MqttLowRequest := TRUE;
	END_IF
END_IF 
                
END_METHOD

METHOD InitMqttDiscoveryAsSwitch
  VAR_INPUT
    Device : POINTER TO FB_PLC_MQTT_DISCOVERY_DEVICE;
    Name : STRING(255);
    DeviceClass : STRING(100) := 'outlet';
    overruleId : STRING(255) := '';
    meta : STRING(255) := '';
  END_VAR
  VAR
    id : STRING(255);
  END_VAR
                  IF InitMqttDone AND NOT initMqttDiscoveryDone THEN
	
	IF CommonTypesAndFunctions.StrEquals(str1:= ADR(overruleId), str2:= ADR('')) THEN
		id := CONCAT(CONCAT(THIS^.DeviceName,'_'), THIS^.InstanceNamePt^); // 'FB_DI_PB_003'
	ELSE
		id := overruleId; // 'MY_PH_GND_HALL_01'
	END_IF
	
	Device^.CreateSwitchEntity(
			Name := name,
			Id := id,
			Meta := meta,
			CommandTopic := THIS^.MQTTSubscribeTopic,
			PayloadOn := 'TRUE',
			PayloadOff := 'FALSE',
			StateTopic := THIS^.MQTTPublishTopic,
			StateOnPayload := 'TRUE',
			StateOffPayload := 'FALSE',
			DeviceClass := DeviceClass);
	
	initMqttDiscoveryDone := TRUE;
END_IF		
                
END_METHOD

METHOD InitMqttDiscoveryAsLight
  VAR_INPUT
    Device : POINTER TO FB_PLC_MQTT_DISCOVERY_DEVICE;
    Name : STRING(255);
    overruleId : STRING(255) := '';
    meta : STRING(255) := '';
  END_VAR
  VAR
    id : STRING(255);
  END_VAR
                  IF InitMqttDone AND NOT initMqttDiscoveryDone THEN
	
	IF CommonTypesAndFunctions.StrEquals(str1:= ADR(overruleId), str2:= ADR('')) THEN
		id := CONCAT(CONCAT(THIS^.DeviceName,'_'), THIS^.InstanceNamePt^); // 'FB_DI_PB_003'
	ELSE
		id := overruleId; // 'MY_PH_GND_HALL_01'
	END_IF
	
	Device^.CreateLightEntity(
			Name := name,
			Id := id,
			Meta := meta,
			CommandTopic := THIS^.MQTTSubscribeTopic,
			PayloadOn := 'TRUE',
			PayloadOff := 'FALSE',
			StateTopic := THIS^.MQTTPublishTopic);

	initMqttDiscoveryDone := TRUE;
END_IF		
                
END_METHOD

METHOD InitMqttDiscoveryAsLock
  VAR_INPUT
    Device : POINTER TO FB_PLC_MQTT_DISCOVERY_DEVICE;
    Name : STRING(255);
    overruleId : STRING(255) := '';
    meta : STRING(255) := '';
  END_VAR
  VAR
    id : STRING(255);
  END_VAR
                  IF InitMqttDone AND NOT initMqttDiscoveryDone THEN
	
	IF CommonTypesAndFunctions.StrEquals(str1:= ADR(overruleId), str2:= ADR('')) THEN
		id := CONCAT(CONCAT(THIS^.DeviceName,'_'), THIS^.InstanceNamePt^); // 'FB_DI_PB_003'
	ELSE
		id := overruleId; // 'MY_PH_GND_HALL_01'
	END_IF
	
	Device^.CreateLockEntity(
		Name := name,
		Id := id,
		Meta := meta,
		CommandTopic := THIS^.MQTTSubscribeTopic,
		PayloadLock := 'TRUE',
		PayloadUnlock := 'FALSE',
		StateTopic := THIS^.MQTTPublishTopic,
		StateUnlocked := 'FALSE',
		StateLocked := 'TRUE');

	initMqttDiscoveryDone := TRUE;
END_IF		
                
END_METHOD

METHOD InitMqttDiscoveryAsSiren
  VAR_INPUT
    Device : POINTER TO FB_PLC_MQTT_DISCOVERY_DEVICE;
    Name : STRING(255);
    overruleId : STRING(255) := '';
    meta : STRING(255) := '';
  END_VAR
  VAR
    id : STRING(255);
  END_VAR
                  IF InitMqttDone AND NOT initMqttDiscoveryDone THEN
	
	IF CommonTypesAndFunctions.StrEquals(str1:= ADR(overruleId), str2:= ADR('')) THEN
		id := CONCAT(CONCAT(THIS^.DeviceName,'_'), THIS^.InstanceNamePt^); // 'FB_DI_PB_003'
	ELSE
		id := overruleId; // 'MY_PH_GND_HALL_01'
	END_IF
	
	Device^.CreateSirenEntity(
			Name := name,
			Id := id,
			Meta := meta,
			CommandTopic := THIS^.MQTTSubscribeTopic,
			PayloadOn := 'TRUE',
			PayloadOff := 'FALSE',
			StateTopic := THIS^.MQTTPublishTopic,
			StateOnPayload := 'TRUE',
			StateOffPayload := 'FALSE');


	initMqttDiscoveryDone := TRUE;
END_IF		
                
END_METHOD
END_FUNCTION_BLOCK

{attribute 'reflection'}
FUNCTION_BLOCK FB_OUTPUT_BISTABLE_MQTT EXTENDS FB_MQTT_BASE IMPLEMENTS MQTT.MQTT_SUBSCRIBE_CALLBACK
  VAR_INPUT
    PRIO_HIGH : BOOL := FALSE;
    PRIO_LOW : BOOL := FALSE;
    TOGGLE : BOOL := FALSE;
    FEEDBACK : BOOL := FALSE;
  END_VAR
  VAR_OUTPUT
    OUT : BOOL;
  END_VAR
  VAR
    {attribute 'instance-path'}
    {attribute 'noinit'}
    InstancePath : STRING;  (* Refelection: object's full instance name *)
    Startup : BOOL := TRUE;
    PreviousFeedback : BOOL;
    HoldTimer : TOF;
    T_hold : TIME := TIME#1s0ms;
    PulseTrigger : BOOL := FALSE;
    MqttDiscoveryMessageLight : MQTT_DISCOVERY_LIGHT;
    MqttDiscoveryMessageLock : MQTT_DISCOVERY_LOCK;
    MqttDiscoveryMessageSiren : MQTT_DISCOVERY_SIREN;
    MqttDiscoveryMessageSwitch : MQTT_DISCOVERY_SWITCH;
  END_VAR

            HoldTimer(PT:= T_hold);

IF PRIO_HIGH THEN
	IF NOT FEEDBACK THEN
		PulseTrigger:=TRUE;
	END_IF
ELSIF(PRIO_LOW AND NOT (PRIO_HIGH)) THEN
	IF FEEDBACK THEN		
		PulseTrigger:=TRUE;
	END_IF
	OUT:= FALSE;
ELSIF MqttHighRequest THEN
	IF NOT FEEDBACK THEN		
		PulseTrigger:=TRUE;
	END_IF
	MqttHighRequest := FALSE;
	MqttLowRequest := FALSE;
ELSIF MqttLowRequest THEN
	IF FEEDBACK THEN		
		PulseTrigger:=TRUE;
	END_IF
	MqttHighRequest := FALSE;
	MqttLowRequest := FALSE;
ELSIF(TOGGLE) THEN	
	PulseTrigger:=TRUE;
END_IF;

IF ((PreviousFeedback <> FEEDBACK) OR Startup) AND InitMqttDone THEN
	pMqttPublishQueue^.AddMessage(
		Payload := BOOL_TO_STRING(FEEDBACK),
		Topic := CONCAT(MqttPublishTopicPrefix^, MqttPublishTopicSuffix),
		Qos := MQTT.QoS.ExactlyOnce,
		MqttRetain := TRUE
	);	
	Startup:=FALSE;
END_IF	

PreviousFeedback := FEEDBACK;
HoldTimer.IN	 := PulseTrigger;
OUT := HoldTimer.Q;

PulseTrigger:=FALSE;
          

METHOD InitMqtt
  VAR_INPUT
    MQTTPublishPrefix : POINTER TO STRING;
    MQTTSubscribePrefix : POINTER TO STRING;
    pMqttPublishQueue : POINTER TO FB_MqttPublishQueue;
    pMqttCallbackCollector : POINTER TO MQTT.CallbackCollector;
  END_VAR
                  SUPER^._InstancePath := THIS^.InstancePath; // Due to reflection its location is important

(*pass trough*)
THIS^.pMqttPublishQueue := pMqttPublishQueue;
THIS^.MqttPublishTopicPrefix:=MQTTPublishPrefix;
THIS^.MQTTSubscribeTopicPrefix:=MQTTSubscribePrefix;
THIS^.pMqttPublishQueue:=pMqttPublishQueue;



SUPER^.InitBaseMqtt();
pMqttCallbackCollector^.put(instance:= THIS^); // register the FB agains the collector so mqtt events can be received


                
END_METHOD

METHOD PublishReceived : BOOL
  VAR_INPUT
    Data : MQTT.CALLBACK_DATA;  (* Collection of recived Data *)
  END_VAR
                  //first check if Mqtt is initialized, otherwise do nothing
IF NOT(InitMqttDone) THEN
	//mark the interface call from the collector as done
	PublishReceived := TRUE;
//check if the packet is for this FB
ELSIF CommonTypesAndFunctions.StrEquals(str1:= ADR(MQTTSubscribeTopic), str2:= Data.TopicOut) THEN
	//mark the interface call from the collector as done
	PublishReceived := TRUE;
	//now process the data
	IF FIND(Data.PayloadString^, 'TRUE') > 0 THEN
		MqttHighRequest := TRUE;
	END_IF
	IF FIND(Data.PayloadString^, 'FALSE') > 0 THEN
		MqttLowRequest := TRUE;
	END_IF
END_IF 
                
END_METHOD

METHOD ConfigureFunctionBlock
  VAR_INPUT
    T_hold : TIME;  (* Default value for click mode, can be overwritten by method call *)
  END_VAR
                  THIS^.T_hold:=T_hold;
                
END_METHOD

METHOD InitMqttDiscoveryAsSwitch
  VAR_INPUT
    Device : POINTER TO FB_PLC_MQTT_DISCOVERY_DEVICE;
    Name : STRING(255);
    DeviceClass : STRING(100) := 'outlet';
    overruleId : STRING(255) := '';
    meta : STRING(255) := '';
  END_VAR
  VAR
    id : STRING(255);
  END_VAR
                  IF InitMqttDone AND NOT initMqttDiscoveryDone THEN
	
	IF CommonTypesAndFunctions.StrEquals(str1:= ADR(overruleId), str2:= ADR('')) THEN
		id := CONCAT(CONCAT(THIS^.DeviceName,'_'), THIS^.InstanceNamePt^); // 'FB_DI_PB_003'
	ELSE
		id := overruleId; // 'MY_PH_GND_HALL_01'
	END_IF
	
	Device^.CreateSwitchEntity(
			Name := name,
			Id := id,
			Meta := meta,
			CommandTopic := THIS^.MQTTSubscribeTopic,
			PayloadOn := 'TRUE',
			PayloadOff := 'FALSE',
			StateTopic := THIS^.MQTTPublishTopic,
			StateOnPayload := 'TRUE',
			StateOffPayload := 'FALSE',
			DeviceClass := DeviceClass);
	
	initMqttDiscoveryDone := TRUE;
END_IF		
                
END_METHOD

METHOD InitMqttDiscoveryAsSiren
  VAR_INPUT
    Device : POINTER TO FB_PLC_MQTT_DISCOVERY_DEVICE;
    Name : STRING(255);
    overruleId : STRING(255) := '';
    meta : STRING(255) := '';
  END_VAR
  VAR
    id : STRING(255);
  END_VAR
                  IF InitMqttDone AND NOT initMqttDiscoveryDone THEN
	
	IF CommonTypesAndFunctions.StrEquals(str1:= ADR(overruleId), str2:= ADR('')) THEN
		id := CONCAT(CONCAT(THIS^.DeviceName,'_'), THIS^.InstanceNamePt^); // 'FB_DI_PB_003'
	ELSE
		id := overruleId; // 'MY_PH_GND_HALL_01'
	END_IF
	
	Device^.CreateSirenEntity(
			Name := name,
			Id := id,
			Meta := meta,
			CommandTopic := THIS^.MQTTSubscribeTopic,
			PayloadOn := 'TRUE',
			PayloadOff := 'FALSE',
			StateTopic := THIS^.MQTTPublishTopic,
			StateOnPayload := 'TRUE',
			StateOffPayload := 'FALSE');

	initMqttDiscoveryDone := TRUE;
END_IF		
                
END_METHOD

METHOD InitMqttDiscoveryAsLock
  VAR_INPUT
    Device : POINTER TO FB_PLC_MQTT_DISCOVERY_DEVICE;
    Name : STRING(255);
    overruleId : STRING(255) := '';
    meta : STRING(255) := '';
  END_VAR
  VAR
    id : STRING(255);
  END_VAR
                  IF InitMqttDone AND NOT initMqttDiscoveryDone THEN
	
	IF CommonTypesAndFunctions.StrEquals(str1:= ADR(overruleId), str2:= ADR('')) THEN
		id := CONCAT(CONCAT(THIS^.DeviceName,'_'), THIS^.InstanceNamePt^); // 'FB_DI_PB_003'
	ELSE
		id := overruleId; // 'MY_PH_GND_HALL_01'
	END_IF
	
	Device^.CreateLockEntity(
		Name := name,
		Id := id,
		Meta := meta,
		CommandTopic := THIS^.MQTTSubscribeTopic,
		PayloadLock := 'TRUE',
		PayloadUnlock := 'FALSE',
		StateTopic := THIS^.MQTTPublishTopic,
		StateUnlocked := 'FALSE',
		StateLocked := 'TRUE');

	initMqttDiscoveryDone := TRUE;
END_IF		
                
END_METHOD

METHOD InitMqttDiscoveryAsLight
  VAR_INPUT
    Device : POINTER TO FB_PLC_MQTT_DISCOVERY_DEVICE;
    Name : STRING(255);
    overruleId : STRING(255) := '';
    meta : STRING(255) := '';
  END_VAR
  VAR
    id : STRING(255);
  END_VAR
                  IF InitMqttDone AND NOT initMqttDiscoveryDone THEN
	
	IF CommonTypesAndFunctions.StrEquals(str1:= ADR(overruleId), str2:= ADR('')) THEN
		id := CONCAT(CONCAT(THIS^.DeviceName,'_'), THIS^.InstanceNamePt^); // 'FB_DI_PB_003'
	ELSE
		id := overruleId; // 'MY_PH_GND_HALL_01'
	END_IF
	
	Device^.CreateLightEntity(
			Name := name,
			Id := id,
			Meta := meta,
			CommandTopic := THIS^.MQTTSubscribeTopic,
			PayloadOn := 'TRUE',
			PayloadOff := 'FALSE',
			StateTopic := THIS^.MQTTPublishTopic);

	initMqttDiscoveryDone := TRUE;
END_IF		
                
END_METHOD
END_FUNCTION_BLOCK

{attribute 'reflection'}
FUNCTION_BLOCK FB_OUTPUT_COVER_MQTT EXTENDS FB_MQTT_BASE IMPLEMENTS MQTT.MQTT_SUBSCRIBE_CALLBACK
  VAR_INPUT
    TOGGLE : BOOL;
    PRIO_LOCK : BOOL;
    PRIO_UP : BOOL;
    PRIO_DN : BOOL;
    {attribute 'input_constant'}
    T_LOCKOUT : TIME := TIME#1s0ms;
    {attribute 'input_constant'}
    T_UD : TIME := TIME#10s0ms;
  END_VAR
  VAR_OUTPUT
    MU : BOOL;
    MD : BOOL;
  END_VAR
  VAR
    {attribute 'instance-path'}
    {attribute 'noinit'}
    InstancePath : STRING;  (* object's full instance name *)
    lock : OSCAT_BASIC.INTERLOCK;
    Cover_State_Timer : TOF;
    internalUp : BOOL;
    internalDown : BOOL;
    MqttRequestStop : BOOL;
    MqttRequestOpen : BOOL;
    MqttRequestClose : BOOL;
    MqttDiscoveryMessage : MQTT_DISCOVERY_COVER;
  END_VAR
  VAR PERSISTENT
    internalDir : BOOL;  (* down = false, up = true *)
  END_VAR

            (* Run the timer to not power the motors for to long *)
Cover_State_Timer(PT:=T_UD);
Cover_State_Timer.IN:=FALSE;

IF NOT(Cover_State_Timer.Q) AND internalUp THEN
	pMqttPublishQueue^.AddMessage(
		Payload := 'OPEN',
		Topic := CONCAT(MqttPublishTopicPrefix^, MqttPublishTopicSuffix),
		Qos := MQTT.QoS.ExactlyOnce,
		MqttRetain := TRUE
	);
END_IF

IF NOT(Cover_State_Timer.Q) AND internalDown THEN
	pMqttPublishQueue^.AddMessage(
		Payload := 'CLOSED',
		Topic := CONCAT(MqttPublishTopicPrefix^, MqttPublishTopicSuffix),
		Qos := MQTT.QoS.ExactlyOnce,
		MqttRetain := TRUE
	);
END_IF


(* Check what to do *)
IF NOT(Cover_State_Timer.Q) AND internalUp THEN // don't run the motors for to long, assume we've reached end and toggle dir
	internalUp := FALSE;
	internalDown := FALSE;
	internalDir := FALSE;
ELSIF NOT(Cover_State_Timer.Q) AND internalDown THEN // don't run the motors for to long, assume we've reached end and toggle dir
	internalUp := FALSE;
	internalDown := FALSE;
	internalDir := TRUE;
ELSIF PRIO_LOCK THEN	
	internalUp := FALSE;
	internalDown := FALSE;
ELSIF PRIO_UP THEN	
	internalUp := TRUE;
	internalDown := FALSE;
	Cover_State_Timer.IN:=TRUE;
ELSIF PRIO_DN THEN	
	internalUp := FALSE;
	internalDown := TRUE;
	Cover_State_Timer.IN:=TRUE;
ELSIF TOGGLE AND (internalUp OR internalDown) THEN	// stop and toggle dir
	internalUp := FALSE;
	internalDown := FALSE;
	internalDir := NOT(internalDir);
ELSIF TOGGLE AND NOT(internalDir) THEN //move down
	internalUp := FALSE;
	internalDown := TRUE;
	Cover_State_Timer.IN:=TRUE;
ELSIF TOGGLE AND internalDir THEN //move upwards
	internalUp := TRUE;
	internalDown := FALSE;	
	Cover_State_Timer.IN:=TRUE;
ELSIF MqttRequestStop THEN
	internalUp := FALSE;
	internalDown := FALSE;
	MqttRequestStop := FALSE;
ELSIF MqttRequestOpen THEN
	internalUp := TRUE;
	internalDown := FALSE;
	MqttRequestOpen := FALSE;
	Cover_State_Timer.IN:=TRUE;;
ELSIF MqttRequestClose THEN
	internalUp := FALSE;
	internalDown := TRUE;
	MqttRequestClose := FALSE;
	Cover_State_Timer.IN:=TRUE;
END_IF

(* make sure only one motor is active at a given time *)
lock(i1 := internalUp, I2 := InternalDown, TL := T_lockout);
MU := lock.Q1;
MD := lock.Q2;
          

METHOD InitMqtt
  VAR_INPUT
    MQTTPublishPrefix : POINTER TO STRING;
    MQTTSubscribePrefix : POINTER TO STRING;
    pMqttPublishQueue : POINTER TO FB_MqttPublishQueue;
    pMqttCallbackCollector : POINTER TO MQTT.CallbackCollector;
  END_VAR
  VAR
    InstanceNamePt : POINTER TO STRING;
  END_VAR
                  SUPER^._InstancePath := THIS^.InstancePath; // Due to reflection its location is important

(*pass trough*)
THIS^.pMqttPublishQueue := pMqttPublishQueue;
THIS^.MqttPublishTopicPrefix:=MQTTPublishPrefix;
THIS^.MQTTSubscribeTopicPrefix:=MQTTSubscribePrefix;
THIS^.pMqttPublishQueue:=pMqttPublishQueue;

SUPER^.InitBaseMqtt();
pMqttCallbackCollector^.put(instance:= THIS^); // register the FB agains the collector so mqtt events can be received
                
END_METHOD

METHOD PublishReceived : BOOL
  VAR_INPUT
    Data : MQTT.CALLBACK_DATA;  (* Collection of recived Data *)
  END_VAR
                  //first check if Mqtt is initialized, otherwise do nothing
IF NOT(InitMqttDone) THEN
	//mark the interface call from the collector as done
	PublishReceived := TRUE;
//check if the packet is for this FB
ELSIF CommonTypesAndFunctions.StrEquals(str1:= ADR(MQTTSubscribeTopic), str2:= Data.TopicOut) THEN
	//mark the interface call from the collector as done
	PublishReceived := TRUE;
	//now process the data
	IF CommonTypesAndFunctions.StrEquals(str1:= Data.PayloadString, str2:= ADR('STOP')) THEN			
		THIS^.MqttRequestStop:=TRUE;
	ELSIF CommonTypesAndFunctions.StrEquals(str1:= Data.PayloadString, str2:= ADR('OPEN')) THEN
		THIS^.MqttRequestOpen:=TRUE;
	ELSIF CommonTypesAndFunctions.StrEquals(str1:= Data.PayloadString, str2:= ADR('CLOSE')) THEN
		THIS^.MqttRequestClose:=TRUE;
	END_IF

END_IF
                
END_METHOD

METHOD ConfigureFunctionBlock : BOOL
  VAR_INPUT
    T_LOCKOUT : TIME;
    T_UD : TIME;
  END_VAR
                  THIS^.T_LOCKOUT:=T_LOCKOUT;
THIS^.T_UD:=T_UD;
                
END_METHOD

METHOD InitMqttDiscovery
  VAR_INPUT
    Device : POINTER TO FB_PLC_MQTT_DISCOVERY_DEVICE;
    Name : STRING(255);
    overruleId : STRING(255) := '';
    meta : STRING(255) := '';
    DeviceClass : STRING(50) := 'shutter';
  END_VAR
  VAR
    id : STRING(255);
  END_VAR
                  IF InitMqttDone AND NOT initMqttDiscoveryDone THEN
	
	IF CommonTypesAndFunctions.StrEquals(str1:= ADR(overruleId), str2:= ADR('')) THEN
		id := CONCAT(CONCAT(THIS^.DeviceName,'_'), THIS^.InstanceNamePt^); // 'FB_DI_PB_003'
	ELSE
		id := overruleId; // 'MY_PH_GND_HALL_01'
	END_IF
	
	Device^.CreateCoverEntity(
		Name := name,
		Id := id,
		Meta := meta,
		CommandTopic := THIS^.MQTTSubscribeTopic,
		PayloadOpen := 'OPEN',
		PayloadClose := 'CLOSE',
		PayloadStop := 'STOP',
		StateTopic := THIS^.MQTTPublishTopic,
		StateOpen := 'OPEN',
		StateClosed := 'CLOSED',
		DeviceClass := DeviceClass
	);

	initMqttDiscoveryDone := TRUE;
END_IF
                
END_METHOD
END_FUNCTION_BLOCK

{attribute 'reflection'}
FUNCTION_BLOCK FB_OUTPUT_DIMMER_MQTT EXTENDS FB_MQTT_BASE IMPLEMENTS MQTT.MQTT_SUBSCRIBE_CALLBACK
  VAR_INPUT
    SINGLE : BOOL;
    LONG : BOOL;
    P_LONG : BOOL;
    PRIO_HIGH : BOOL := FALSE;
    PRIO_LOW : BOOL := FALSE;
    SET : BOOL;
    VAL : BYTE;
    RST : BOOL;
  END_VAR
  VAR_OUTPUT
    Q : BOOL;
    Q_OUT : WORD;
    OUT : WORD;
  END_VAR
  VAR
    {attribute 'instance-path'}
    {attribute 'noinit'}
    InstancePath : STRING;  (* Refelection: object's full instance name *)
    t3 : OSCAT_BASIC.TON;
    dim : OSCAT_BASIC._RMP_B;
    dir : BOOL;
    OUT_Internal : BYTE;
    LIN_TRAFO : Util.LIN_TRAFO;
    enabled : BOOL := TRUE;
    Startup : BOOL := TRUE;
    OutputDimmer : BOOL;
    Qos_Dimm : MQTT.QoS;
    Delta_Dimm : INT;
    T_Debounce : TIME := TIME#10ms;  (* Default values for dimmer, can be overwritten by method call *)
    T_Reconfig : TIME := TIME#10s0ms;
    T_On_Max : TIME := TIME#0ms;
    T_Dimm_Start : TIME := TIME#400ms;
    T_Dimm : TIME := TIME#1s0ms;
    Min_On : BYTE := 100;
    Max_On : BYTE := 200;
    Soft_Dimm : BOOL := TRUE;
    Rst_Out : BOOL := FALSE;
    OUT_LinearScaleMin : INT := 10000;
    OUT_LinearScaleMax : INT := 32767;
    DmxChannel : INT;  (* DMX specific *)
    DmxWidth : INT;
    DmxUniverse : INT;
    pDmxValues : POINTER TO oscat_network.NETWORK_BUFFER_SHORT;
    InitDmxDone : BOOL := FALSE;
    OUT_Target : BYTE;
    SoftDimToValue : BOOL;
    SoftDimToQFalse : BOOL;
    UpdateValueStep : BYTE := 4;
    OUT_Internal_tmp : BYTE;
    curve : DINT := DIMMER_CURVE.linear;
    wait : TON;
    Step : INT := 0;
    dimmedValue : INT := 1;
    waitTimeAtTop : TIME := TIME#200ms;  (* one time before and after blink *)
    blinkValue : BYTE := 100;
    blinkEnabled : BOOL := FALSE;
    MqttDiscoveryMessage : MQTT_DISCOVERY_LIGHT_DIMMER;
  END_VAR
  VAR PERSISTENT
    PreviousOUT : BYTE;  (* To retain output state through powercycles *)
    PreviousQ : BOOL;  (* To retain output state through powercycles *)
  END_VAR

            

IF Startup THEN
	OUT := PreviousOUT;
	Q := PreviousQ;
END_IF

IF RST THEN
	IF rst_out THEN OUT_Internal := 0; END_IF;
	Q := FALSE;
	dir := OUT_Internal > 127;
ELSIF PRIO_HIGH THEN
	Q := TRUE;
	OUT_Internal := 255;
ELSIF PRIO_LOW THEN
	Q := FALSE;
ELSIF MqttHighRequest THEN
	Q:= TRUE;
	MqttHighRequest := FALSE;
	MqttLowRequest := FALSE;
ELSIF MqttLowRequest THEN
	Q:= FALSE;
	MqttHighRequest := FALSE;
	MqttLowRequest := FALSE;
ELSIF set THEN
	OUT_Internal := val;
	Q := TRUE;
	(* set direction to up when value < 127 otherwise set dir down dir is reversed because next action will reverse again *)
	dir := OUT_Internal > 127;
ELSIF SINGLE THEN
	(* a single click reverses output Q *)
	Q := NOT Q;
	(* when dimmer is turned on we need to limit out to min and max limits *)
	IF Q THEN OUT_Internal := LIMIT(MAX(OUT_Internal,1), OUT_Internal, MAX_ON);	END_IF;
	(* set the appropriate direction of dimmer dir is reversed because next action will reverse again *)
	dir := OUT_Internal > 127;
ELSIF LONG THEN
	IF NOT Q THEN
		IF SOFT_DIMM THEN
			OUT_Internal := 1;
			dir := TRUE;
		ELSE
			OUT_Internal := LIMIT(MAX(MIN_ON,1), OUT_Internal, MAX_ON);
			DIR := OUT_Internal < 127;
		END_IF;
		Q := TRUE;
	ELSE
		(* reverse direction with every long click *)
		dir := NOT dir;
	END_IF;
END_IF;


(* while dimming is active ramp the output out up or down *)
dim(DIR := dir, e := P_LONG AND Q, TR := T_DIMM, rmp := OUT_Internal);

(* reverse direction when limits are reached *)
IF OUT_Internal = 0 THEN
	dir := TRUE;
ELSIF OUT_Internal = 255 THEN
	dir := FALSE;
END_IF;

(* limit the maximum runtime *)
IF t_ON_MAX > t#0s THEN
	t3(in := q, pt := T_ON_MAX);
	Q := Q XOR t3.Q;
END_IF;

(* Scale the internal OUT to the actual OUT *)
LIN_TRAFO(
		IN:= OUT_Internal,
		IN_MIN:= 0,
		IN_MAX:= 255,
		OUT_MIN:=OUT_LinearScaleMin,
		OUT_MAX:=OUT_LinearScaleMax
	);
OUT:= REAL_TO_WORD(LIN_TRAFO.OUT);
IF Q THEN
	Q_OUT:= OUT;
ELSE
	Q_OUT:= 0;
END_IF

IF ((ABS(BYTE_TO_INT(PreviousOUT) - BYTE_TO_INT(OUT_Internal)) >= Delta_Dimm) OR Startup AND OUT_Internal <> PreviousOUT OR Startup AND OutputDimmer) AND InitMqttDone THEN
	PreviousOUT:=OUT_Internal;
	pMqttPublishQueue^.AddMessage(		
		Payload := BYTE_TO_STRING(OUT_Internal),
		Topic := CONCAT(THIS^.MQTTPublishTopic,'/OUT'),
		Qos := MQTT.QoS.ExactlyOnce,
		MqttRetain := TRUE
	);
END_IF

IF (Q <> PreviousQ OR Startup) AND InitMqttDone THEN
	PreviousQ:=Q;
	pMqttPublishQueue^.AddMessage(
		Payload := BOOL_TO_STRING(Q),
		Topic := CONCAT(THIS^.MQTTPublishTopic,'/Q'),
		Qos := Qos_Dimm,
		MqttRetain := TRUE
	);
END_IF

Startup:=FALSE;

(* DMX specific *)
IF InitDmxDone THEN 
	IF Q THEN
		IF pDmxValues^.BUFFER[DmxChannel-1] <> OUT_Internal THEN
			pDmxValues^.BUFFER[DmxChannel-1] := OUT_Internal;
		END_IF
	ELSE 
		IF pDmxValues^.BUFFER[DmxChannel-1] <> 0 THEN
			pDmxValues^.BUFFER[DmxChannel-1] := 0;
		END_IF
	END_IF
END_IF
IF SoftDimToValue AND OUT_Internal = OUT_Target THEN // If the same, softdim to value is done
	SoftDimToValue := FALSE;
	IF SoftDimToQFalse THEN
		SoftDimToQFalse := FALSE;
		OUT_Internal := OUT_Internal_tmp;
		PreviousOUT:=OUT_Internal;
	END_IF
END_IF
Startup:=FALSE;

(* DMX specific *)

          

METHOD PublishReceived : BOOL
  VAR_INPUT
    Data : MQTT.CALLBACK_DATA;  (* Collection of recived Data *)
  END_VAR
                  //first check if Mqtt is initialized, otherwise do nothing
IF NOT(InitMqttDone) THEN
	//mark the interface call from the collector as done
	PublishReceived := TRUE;
//check if the packet is for this FB
ELSIF CONCAT(MQTTSubscribeTopic,'/Q') =  Data.TopicOut^ THEN
	IF CommonTypesAndFunctions.StrEquals(str1:= Data.PayloadString, str2:= ADR('TRUE')) THEN
		MqttHighRequest := TRUE;
	ELSIF CommonTypesAndFunctions.StrEquals(str1:= Data.PayloadString, str2:= ADR('FALSE')) THEN
		MqttLowRequest := TRUE;
	END_IF;
	
ELSIF CONCAT(MQTTSubscribeTopic,'/OUT') =  Data.TopicOut^ THEN
	IF OSCAT_BASIC.IS_CC(str:= Data.PayloadString^,cmp:='0123456789.') AND THIS^.PRIO_HIGH = FALSE THEN
		THIS^.OUT_Target:=STRING_TO_BYTE(Data.PayloadString^);
		THIS^.SoftDimToValue:=TRUE;
	END_IF
	
	
// Legacy! backwards compatiably with /+ topics instead of /#
ELSIF CommonTypesAndFunctions.StrEqualsAtStart(str1:= ADR(MQTTSubscribeTopic), str2:= Data.TopicOut) THEN
	//mark the interface call from the collector as done
	PublishReceived := TRUE;
	//now process the data
	IF CommonTypesAndFunctions.StrEquals(str1:= Data.PayloadString, str2:= ADR('TRUE')) THEN
		MqttHighRequest := TRUE;
	ELSIF CommonTypesAndFunctions.StrEquals(str1:= Data.PayloadString, str2:= ADR('FALSE')) THEN
		MqttLowRequest := TRUE;
	ELSIF OSCAT_BASIC.IS_CC(str:= Data.PayloadString^,cmp:='0123456789.') AND THIS^.PRIO_HIGH = FALSE THEN
		THIS^.OUT_Target:=STRING_TO_BYTE(Data.PayloadString^);
		THIS^.SoftDimToValue:=TRUE;
	END_IF
END_IF 
                
END_METHOD

METHOD ConfigureFunctionBlock
  VAR_INPUT
    T_Debounce : TIME := TIME#10ms;  (* Default values for dimmer, can be overwritten by method call *)
    T_Reconfig : TIME := TIME#10s0ms;
    T_On_Max : TIME := TIME#0ms;
    T_Dimm_Start : TIME := TIME#400ms;
    T_Dimm : TIME := TIME#3s0ms;
    Min_On : BYTE := 50;
    Max_On : BYTE := 255;
    Soft_Dimm : BOOL := TRUE;
    Rst_Out : BOOL := FALSE;
    OUT_LinearScaleMin : INT := 0;
    OUT_LinearScaleMax : INT := 32767;
  END_VAR
                  THIS^.T_Debounce:=T_Debounce;
THIS^.T_Reconfig:=T_Reconfig;
THIS^.T_On_Max:=T_On_Max;
THIS^.T_Dimm_Start:=T_Dimm_Start;
THIS^.T_Dimm:=T_Dimm;
THIS^.Min_On:=Min_On;
THIS^.Max_On:=Max_On;
THIS^.Soft_Dimm:=Soft_Dimm;
THIS^.Rst_Out:=Rst_Out;
THIS^.OUT_LinearScaleMin:=OUT_LinearScaleMin;
THIS^.OUT_LinearScaleMax:=OUT_LinearScaleMax;
                
END_METHOD

METHOD InitMqtt
  VAR_INPUT
    MQTTPublishPrefix : POINTER TO STRING;
    MQTTSubscribePrefix : POINTER TO STRING;
    pMqttPublishQueue : POINTER TO FB_MqttPublishQueue;
    pMqttCallbackCollector : POINTER TO MQTT.CallbackCollector;
    OutputDimmer : BOOL;  (* Dimmer specific *)
    Qos_Dimm : MQTT.QoS;
    Delta_Dimm : INT;
  END_VAR
                  SUPER^._InstancePath := THIS^.InstancePath; // Due to reflection its location is important

(*pass trough*)
THIS^.pMqttPublishQueue := pMqttPublishQueue;
THIS^.MqttPublishTopicPrefix:=MQTTPublishPrefix;
THIS^.MQTTSubscribeTopicPrefix:=MQTTSubscribePrefix;
THIS^.pMqttPublishQueue:=pMqttPublishQueue;

// Dimmer specific
THIS^.OutputDimmer:=OutputDimmer;
THIS^.Qos_Dimm:=Qos_Dimm;
THIS^.Delta_Dimm:=Delta_Dimm;


SUPER^.InitBaseMqtt();
pMqttCallbackCollector^.put(instance:= THIS^); // register the FB agains the collector so mqtt events can be received


                
END_METHOD

METHOD initDMX
  VAR_INPUT
    DmxChannel : INT;
    DmxWidth : INT := 1;
    DmxUniverse : INT := 1;
    pDmxValues : POINTER TO oscat_network.NETWORK_BUFFER_SHORT;
  END_VAR
                  
IF NOT THIS^.InitDmxDone THEN
	THIS^.DmxChannel := DmxChannel;
	THIS^.pDmxValues := pDmxValues;
	THIS^.DmxWidth := DmxWidth;
	THIS^.InitDmxDone := TRUE;
	
	THIS^.InitDmxDone := TRUE;
END_IF
                
END_METHOD

METHOD InitMqttDiscovery
  VAR_INPUT
    Device : POINTER TO FB_PLC_MQTT_DISCOVERY_DEVICE;
    Name : STRING(255);
    overruleId : STRING(255) := '';
    meta : STRING(255) := '';
  END_VAR
  VAR
    id : STRING(255);
  END_VAR
                  IF InitMqttDone AND NOT initMqttDiscoveryDone THEN
	
	IF CommonTypesAndFunctions.StrEquals(str1:= ADR(overruleId), str2:= ADR('')) THEN
		id := CONCAT(CONCAT(THIS^.DeviceName,'_'), THIS^.InstanceNamePt^); // 'FB_DI_PB_003'
	ELSE
		id := overruleId; // 'MY_PH_GND_HALL_01'
	END_IF
	
	Device^.CreateLightDimmerEntity(
		Name := name,
		Id := Id,
		Meta := meta,
		CommandTopic := CONCAT(THIS^.MQTTSubscribeTopic,'/Q'),
		PayloadOn := 'TRUE',
		PayloadOff := 'FALSE',
		StateTopic := CONCAT(THIS^.MQTTPublishTopic,'/Q'),
		BrightnessCommandTopic := CONCAT(THIS^.MQTTSubscribeTopic,'/OUT'),
		BrightnessStateTopic := CONCAT(THIS^.MQTTPublishTopic,'/OUT'),
		BrightnessScale := 255,
		DmxChannel := THIS^.DmxChannel,
		DmxWidth := THIS^.DmxWidth,
		DmxUniverse := THIS^.DmxUniverse);

	initMqttDiscoveryDone := TRUE;
END_IF
                
END_METHOD
END_FUNCTION_BLOCK

{attribute 'reflection'}
FUNCTION_BLOCK FB_PLC_MQTT_DISCOVERY_DEVICE EXTENDS FB_BASE_MQTT_DISCOVERY_DEVICE

            
          

METHOD initPlcDevice
  VAR_INPUT
    url : STRING := '';
    availabilityTopic : STRING;
    availabilityOnline : STRING;
    availabilityOffline : STRING;
    MqttDiscoveryPrefix : STRING;
    pMqttPublishQueue : POINTER TO FB_MqttPublishQueue;
  END_VAR
  VAR
    Author : STRING;
    LocalUrl : STRING;
    iSplitLocation : INT;
    AdapterInfo : SOCK_ADAPTER_INFORMATION;
    hAdapter : RTS_IEC_HANDLE;
    udiStructSize : UDINT := SIZEOF(AdapterInfo);
    rResult : RTS_IEC_RESULT;
    sIpAddr : STRING(15);
    sMacAddr : STRING(17);
    xFirstAdapter : BOOL;
    xReadInfo : BOOL;
    xRead : BOOL;
    iecResult : SysTypes.RTS_IEC_RESULT;
    dwType : DWORD;
    dwTargetId : DWORD;
    wsDeviceName : WSTRING;
    wsDev : DINT := SIZEOF(wsDeviceName);
    udiProcessorId : UDINT;
    udiOsId : UDINT;
    sSerialNumber : STRING;
    psSerialNumber : POINTER TO STRING := ADR(sSerialNumber);
    diSerialNumber : DINT := SIZEOF(sSerialNumber);
    xInit : BOOL := TRUE;
  END_VAR
                  IF xInit THEN
    xInit := FALSE;
	
    xFirstAdapter := TRUE;
    rResult := 0;
    WHILE rResult = 0 DO   
        IF xFirstAdapter THEN
            hAdapter := SysSockGetFirstAdapterInfo(ADR(AdapterInfo), ADR(udiStructSize), ADR(rResult));
        ELSE   
            hAdapter := SysSockGetNextAdapterInfo(hAdapter, ADR(AdapterInfo), ADR(udiStructSize), ADR(rResult));
        END_IF
        IF rResult = 0 THEN
            sIpAddr := Standard.CONCAT(BYTE_TO_STRING(AdapterInfo.IpAddr.S_un_b.s_b1),'.');
            sIpAddr := Standard.CONCAT(sIpAddr,BYTE_TO_STRING(AdapterInfo.IpAddr.S_un_b.s_b2));
            sIpAddr := Standard.CONCAT(sIpAddr,'.');
            sIpAddr := Standard.CONCAT(sIpAddr,BYTE_TO_STRING(AdapterInfo.IpAddr.S_un_b.s_b3));
            sIpAddr := Standard.CONCAT(sIpAddr,'.');
            sIpAddr := Standard.CONCAT(sIpAddr,BYTE_TO_STRING(AdapterInfo.IpAddr.S_un_b.s_b4));
            sMacAddr := Standard.CONCAT(SM0.Byte_To_HexString(AdapterInfo.abyMac[0]),'-');
            sMacAddr := Standard.CONCAT(sMacAddr,SM0.Byte_To_HexString(AdapterInfo.abyMac[1]));
            sMacAddr := Standard.CONCAT(sMacAddr,'-');
            sMacAddr := Standard.CONCAT(sMacAddr,SM0.Byte_To_HexString(AdapterInfo.abyMac[2]));
            sMacAddr := Standard.CONCAT(sMacAddr,'-');
            sMacAddr := Standard.CONCAT(sMacAddr,SM0.Byte_To_HexString(AdapterInfo.abyMac[3]));
            sMacAddr := Standard.CONCAT(sMacAddr,'-');
            sMacAddr := Standard.CONCAT(sMacAddr,SM0.Byte_To_HexString(AdapterInfo.abyMac[4]));
            sMacAddr := Standard.CONCAT(sMacAddr,'-');
            sMacAddr := Standard.CONCAT(sMacAddr,SM0.Byte_To_HexString(AdapterInfo.abyMac[5]));
        END_IF
        xFirstAdapter := FALSE;   
    END_WHILE


 
    //  Control WinV3: 4096 - 0000 0001
    iecResult := SysTarget.SysTargetGetType(pulType := ADR(dwType));
    iecResult := SysTarget.SysTargetGetId(pulTargetId := ADR(dwTargetId));
 
    iecResult := SysTarget.SysTargetGetDeviceName(pwszName := ADR(wsDeviceName), pnMaxLength := ADR(wsDev));
 
 
    //Unique RT identifier
    iecResult := SysTarget.SysTargetGetSerialNumber(ppsSerialNumber := ADR(psSerialNumber), pnMaxLen := ADR(diSerialNumber));

	
    pApp := AppFindApplicationByName(pszString := sAppName, pResult := ADR(iecResult));   
    pstAppInfo := AppGetApplicationInfo(pApp := pApp, pResult := ADR(iecResult));   
		//         MqttVariables.version := pstAppInfo^.pstVersion^;
		//         MqttVariables.desc := pstAppInfo^.pstDescription^;

    IF iecResult = 0 THEN
		
		iSplitLocation := COL.Stu.StrFindA(
			pst1:= ADR(THIS^.InstanceName), 
			pst2:= ADR('.'), 
			uiSearchStart:= 1
		) - 1;
	
	
		IF CommonTypesAndFunctions.StrEquals(str1:= ADR(pstAppInfo^.pstAuthor), str2:= ADR('')) THEN
			Author := 'MichielVanwelsenaere et al.';
		ELSE
			Author := pstAppInfo^.pstAuthor^; // 'DIMMER_GND_HALL_01'
		END_IF	
		
		IF CommonTypesAndFunctions.StrEquals(ADR(url), ADR('')) THEN
			LocalUrl := CONCAT('https://', sIpAddr);
		ELSE
			LocalUrl := url;
		END_IF
			
		SUPER^.initBaseDevice(
			Name := LEFT(THIS^.InstanceName,iSplitLocation),
			ConfigurationUrl := LocalUrl,
			Identifiers := psSerialNumber^,
			Manufacturer := Author,
			Model := pstAppInfo^.pstDescription^,
			SoftwareVersion := CONCAT(CONCAT( DT_TO_STRING(pstAppInfo^.dtLastChanges),' '), pstAppInfo^.pstProjectName^),
			HardwareVersion := WSTRING_TO_STRING(wsDeviceName),
			IpAddress := sIpAddr,
			MacAddress := sMacAddr,
			availabilityTopic := availabilityTopic,			
			availabilityOnline := availabilityOnline,
			availabilityOffline := availabilityOffline,
			MqttDiscoveryPrefix := MqttDiscoveryPrefix,
			pMqttPublishQueue := pMqttPublishQueue);
    END_IF
END_IF




                
END_METHOD
END_FUNCTION_BLOCK

FUNCTION_BLOCK FB_RS485_BUSCONTROLLER
  VAR_OUTPUT
    BusOcupied : BOOL := TRUE;  (* Set this to True by default at startup to allow for some RS485 devices to boot up at power interuptions *)
  END_VAR
  VAR
    StartupDelay : TIME := TIME#5s0ms;  (* Amount of time that should be waited on PLC startup to start using the RS485 bus *)
    SilenceTime : TIME := TIME#20ms;  (* This is the silence time between two requests *)
    Startup : BOOL := TRUE;  (* Used to detect startup *)
    tonDelay : TON;  (* To manage silence time and startup delay *)
    devices : ARRAY[0..31] OF RS485Device;  (* collection of devices on the bus *)
    devicesCount : INT := 0;  (* total number of devices registred on the bus *)
    selectedDevice : INT := 0;  (* index of the active device on the bus *)
    deviceActive : BOOL;
    loopCounter : INT;
    ActiveRtuQuery : RS485_RtuQuery;
    BusTrigger : POINTER TO BOOL;
    QueryReady : Standard.F_TRIG;
    BusData : POINTER TO ARRAY[0..124] OF WORD;
    BusError : POINTER TO BOOL;
    exc : __SYSTEM.ExceptionCode;
  END_VAR

            IF Startup THEN
	tonDelay.PT := StartupDelay;
	tonDelay.IN := TRUE;
	Startup := FALSE;
END_IF

QueryReady(CLK := BusTrigger^);
BusOcupied := NOT(tonDelay.Q);
tonDelay();

// check if there's a device that requires bus time and if so, launch the query
IF busOcupied = FALSE AND deviceActive = FALSE AND devicesCount <> 0 AND NOT QueryReady.Q THEN
	FOR loopCounter := 0 TO devicesCount - 1 DO
		IF deviceActive = FALSE AND devices[loopCounter].RequestBusTime() THEN
			selectedDevice := loopCounter;
			THIS^.SetBusOccupied();
			ActiveRtuQuery := devices[selectedDevice].GetRtuQuery();
			BusTrigger^ := TRUE;
			EXIT;
		END_IF
	END_FOR;
END_IF

//watch the trigger, when completed call the FB with the data, release the bus
IF QueryReady.Q THEN
	devices[selectedDevice].ProcessDataArray(BusError, BusData);
	THIS^.ReleaseBus();
END_IF


//let the busdevices to their work
//FOR loopCounter := 0 TO devicesCount - 1 DO
//	devices[loopCounter]();
// END_FOR;
          

METHOD RegisterDevice
  VAR_INPUT
    device : RS485Device;
  END_VAR
                  IF devicesCount <> 32 THEN
	devices[devicesCount] := device;
	devicesCount := devicesCount + 1;
END_IF
                
END_METHOD

METHOD ReleaseBus
                  // Start a timer to release the bus
THIS^.tonDelay.PT := THIS^.SilenceTime;
THIS^.tonDelay.IN := TRUE;
THIS^.deviceActive := FALSE;
                
END_METHOD

METHOD SetBusOccupied
                  THIS^.tonDelay.IN := FALSE;
THIS^.deviceActive := TRUE;
                
END_METHOD

METHOD Init
  VAR_INPUT
    StartupDelay : TIME;  (* Amount of time that should be waited on PLC startup to start using the RS485 bus, can prevent errors due to devices not booted up yet *)
    SilenceTime : TIME;  (* This is the silence time between two requests *)
    BusTrigger : POINTER TO BOOL;  (* pointer to the bool that controls triggering busrequests *)
    BusData : POINTER TO ARRAY[0..124] OF WORD;
    BusError : POINTER TO BOOL;
  END_VAR
                  THIS^.StartupDelay := StartupDelay;
THIS^.SilenceTime := SilenceTime;
THIS^.BusTrigger := BusTrigger;
THIS^.BusData := BusData;
THIS^.BusError := BusError;
                
END_METHOD
END_FUNCTION_BLOCK

{attribute 'reflection'}
FUNCTION_BLOCK FB_RS485_DUCO_DUCOBOX_MQTT IMPLEMENTS RS485Device, MQTT.MQTT_SUBSCRIBE_CALLBACK
  VAR_OUTPUT
    ACTIVEPOWER : REAL := 0;
    DataAvailable : BOOL := FALSE;
    Error : BOOL := FALSE;
  END_VAR
  VAR
    {attribute 'instance-path'}
    {attribute 'noinit'}
    InstanceName : STRING;  (* object's full instance name *)
    Startup : BOOL := TRUE;
    InitMqttDone : BOOL;
    MqttPublishTopicPrefix : POINTER TO STRING;
    MqttPublishTopicSuffix : STRING(50);
    MQTTSubscribeTopic : STRING(50);
    pMqttPublishQueue : POINTER TO FB_MqttPublishQueue;
    InitRS485Done : BOOL := FALSE;
    timerData : TON;
    isDataUpdated : BOOL := FALSE;
    Nodes : ARRAY[2..30] OF FB_RS485_DUCO_DUCOBOX_NODE_MQTT;
    NodePointer : UINT := 2;
    ActiveNode : INT := 0;
    loopCounter : INT;
    ReadMasterUnitQuery : RS485_RtuQuery := (FunctionCode := 4, ReadAddress := 10, ReadQuantity := 6);
    WriteQueryReady : BOOL := FALSE;
    WriteQueryBeingExecuted : BOOL := FALSE;
    WriteQuerySuffix : STRING;
    WriteQueryPayload : STRING;
    WriteQuery : RS485_RtuQuery := (FunctionCode := 6, WriteQuantity := 1);
  END_VAR

            timerData();

FOR loopCounter := 2 TO 30 DO
	Nodes[loopCounter]();
END_FOR
          

METHOD ProcessDataArray
  VAR_INPUT
    Error : POINTER TO BOOL;
    Data : POINTER TO ARRAY[0..124] OF WORD;
  END_VAR
                  THIS^.Error := Error^;

IF Error^ AND NOT WriteQueryBeingExecuted THEN
	PubMqttMessage(Suffix := '/availability', Data := 'offline');
ELSE
	PubMqttMessage(Suffix := '/availability', Data := 'online');
END_IF

IF WriteQueryBeingExecuted THEN
	WriteQueryReady := FALSE;
	WriteQueryBeingExecuted := FALSE;
	IF NOT Error^ THEN
		PubMqttMessage(Suffix := CONCAT('/', WriteQuerySuffix), Data := WriteQueryPayload);
	END_IF
// data for master unit (= main node)
ELSIF THIS^.ActiveNode = 1 THEN
	THIS^.timerData.IN := TRUE;
	THIS^.ActiveNode := 0;
	
	IF NOT Error^ THEN
 		PubMqttMessage(Suffix := '/1/read/0', Data := WORD_TO_STRING(Data^[0]));
 		PubMqttMessage(Suffix := '/1/read/1', Data := WORD_TO_STRING(Data^[1]));
 		PubMqttMessage(Suffix := '/1/read/2', Data := WORD_TO_STRING(Data^[2]));
 		PubMqttMessage(Suffix := '/1/read/3', Data := WORD_TO_STRING(Data^[3]));
 		PubMqttMessage(Suffix := '/1/read/4', Data := WORD_TO_STRING(Data^[4]));
 		PubMqttMessage(Suffix := '/1/read/5', Data := WORD_TO_STRING(Data^[5]));
	END_IF
// data for nodes
ELSIF THIS^.ActiveNode > 1 THEN	
	THIS^.Nodes[ActiveNode].ProcessDataArray(
		Data := Data,
		Error := Error
	);
	THIS^.ActiveNode := 0;
END_IF
                
END_METHOD

METHOD InitRS485
  VAR_INPUT
    DataPollingInterval : TIME;
    DeviceAddress : BYTE;
  END_VAR
                  THIS^.timerData.PT := DataPollingInterval;
THIS^.ReadMasterUnitQuery.DeviceId := DeviceAddress;
THIS^.WriteQuery.DeviceId := DeviceAddress;
THIS^.timerData.IN := TRUE;

THIS^.InitRS485Done := TRUE;
                
END_METHOD

METHOD InitMqtt
  VAR_INPUT
    MQTTPublishPrefix : POINTER TO STRING;
    MQTTSubscribePrefix : POINTER TO STRING;
    pMqttPublishQueue : POINTER TO FB_MqttPublishQueue;
    pMqttCallbackCollector : POINTER TO MQTT.CallbackCollector;
  END_VAR
  VAR
    InstanceNamePt : POINTER TO STRING;
  END_VAR
                  THIS^.pMqttPublishQueue := pMqttPublishQueue;
THIS^.MqttPublishTopicPrefix := MQTTPublishPrefix;

InstanceNamePt := CommonTypesAndFunctions.FindLastDot(ADR(THIS^.InstanceName)) + 1;
THIS^.MqttPublishTopicSuffix := InstanceNamePt^;
THIS^.MQTTSubscribeTopic := CONCAT(MQTTSubscribePrefix^ ,THIS^.MqttPublishTopicSuffix);

// register the FB agains the collector so mqtt events can be received
pMqttCallbackCollector^.put(instance:= THIS^);


FOR loopCounter := 2 TO 30 DO
		Nodes[loopCounter].InitMqtt(
			MQTTPublishPrefix := MQTTPublishPrefix,
			MqttPublishTopicSuffix := InstanceNamePt^,
			pMqttPublishQueue := pMqttPublishQueue
		);
END_FOR

InitMqttDone := TRUE;
                
END_METHOD

METHOD RequestBusTime : BOOL
                  IF NOT InitRS485Done THEN	
	RequestBusTime := FALSE;
ELSIF WriteQueryReady THEN
	RequestBusTime := TRUE;	
ELSIF timerData.Q THEN // Master node
	RequestBusTime := TRUE;
	THIS^.ActiveNode := 1;
ELSIF NodePointer > 2 THEN// other nodes, if configured
	FOR loopCounter := 2 TO 30 DO
		IF Nodes[loopCounter].RequestBusTime() AND RequestBusTime = FALSE THEN
			THIS^.ActiveNode := loopCounter;
			RequestBusTime := TRUE;	
		END_IF
	END_FOR
ELSE
	RequestBusTime := FALSE;
END_IF

                
END_METHOD

METHOD GetRtuQuery : RS485_RtuQuery
                  IF WriteQueryReady THEN
	GetRtuQuery := THIS^.WriteQuery;
	WriteQueryBeingExecuted := TRUE;
// master
ELSIF ActiveNode = 1 THEN
	THIS^.timerData.IN := FALSE;
	GetRtuQuery := THIS^.ReadMasterUnitQuery;
// other nodes
ELSIF ActiveNode > 1 THEN
	GetRtuQuery := THIS^.Nodes[ActiveNode].GetRtuQuery();	
END_IF
                
END_METHOD

METHOD PubMqttMessage
  VAR_INPUT
    Suffix : STRING(100);
    Data : STRING(100);
  END_VAR
                  IF InitMqttDone THEN
		pMqttPublishQueue^.AddMessage(
			Payload := Data,
			Topic := CONCAT(CONCAT(MqttPublishTopicPrefix^, MqttPublishTopicSuffix), Suffix ),
			Qos := MQTT.QoS.ExactlyOnce,
			MqttRetain := FALSE
		);
END_IF
                
END_METHOD

METHOD PublishReceived : BOOL
  VAR_INPUT
    Data : MQTT.CALLBACK_DATA;  (* Collection of recived Data *)
  END_VAR
  VAR
    SubTopic : STRING;
    NodeNumber : STRING;
    NodeRegister : STRING;
  END_VAR
                  //first check if Mqtt is initialized, otherwise do nothing
IF NOT(InitMqttDone) THEN
	//mark the interface call from the collector as done
	PublishReceived := TRUE;
//check if the packet is for this FB
ELSIF MQTTSubscribeTopic = LEFT(Data.TopicOut^, LEN(MQTTSubscribeTopic)) THEN
	//mark the interface call from the collector as done
	PublishReceived := TRUE;
	// process the data
	SubTopic := RIGHT(Data.TopicOut^, 9); // 2/write/9 -> 10 chars
	NodeNumber := LEFT(SubTopic, 1);
	NodeRegister := RIGHT(SubTopic, 1);
	
	IF FIND(SubTopic, 'write') > 0 AND
		OSCAT_BASIC.IS_NUM(NodeNumber) AND
		OSCAT_BASIC.IS_NUM(NodeRegister) AND
		OSCAT_BASIC.IS_NUM(Data.PayloadString^) THEN
			WriteQuery.WriteAddress := (STRING_TO_UINT(NodeNumber) * 10) + STRING_TO_UINT(NodeRegister);
			WriteQuery.WriteData[0] := STRING_TO_WORD(Data.PayloadString^);
			WriteQuerySuffix := SubTopic;
			WriteQueryPayload := Data.PayloadString^;
			WriteQueryReady := TRUE;
	END_IF
END_IF
                
END_METHOD

METHOD AddNode : BOOL
  VAR_INPUT
    DataPollingInterval : TIME;
  END_VAR
                  THIS^.Nodes[NodePointer].InitNode(
	DeviceAddress := THIS^.ReadMasterUnitQuery.DeviceId,
	NodeNumber := NodePointer -1,
	DataPollingInterval := DataPollingInterval
);

NodePointer := NodePointer + 1;
                
END_METHOD
END_FUNCTION_BLOCK

FUNCTION_BLOCK FB_RS485_DUCO_DUCOBOX_NODE_MQTT
  VAR
    NodeNumber : UINT;
    InitMqttDone : BOOL;
    MqttPublishTopicPrefix : POINTER TO STRING;
    MqttPublishTopicSuffix : STRING(51);
    pMqttPublishQueue : POINTER TO FB_MqttPublishQueue;
    NodeInitialized : BOOL := FALSE;
    timerData : TON;
    RtuQueryRead : RS485_RtuQuery := (FunctionCode := 4, ReadAddress := 20, ReadQuantity := 6);
  END_VAR

            timerData();


          

METHOD GetRtuQuery : RS485_RtuQuery
                  IF timerData.Q THEN
	THIS^.timerData.IN := FALSE;
	GetRtuQuery := THIS^.RtuQueryRead;	
END_IF
                
END_METHOD

METHOD ProcessDataArray
  VAR_INPUT
    Error : POINTER TO BOOL;
    Data : POINTER TO ARRAY[0..124] OF WORD;
  END_VAR
                  THIS^.timerData.IN := TRUE;

IF NOT Error^ THEN
	PubMqttMessage(Suffix := '/read/0', Data := WORD_TO_STRING(Data^[0]));
	PubMqttMessage(Suffix := '/read/1', Data := WORD_TO_STRING(Data^[1]));
	PubMqttMessage(Suffix := '/read/2', Data := WORD_TO_STRING(Data^[2]));
	PubMqttMessage(Suffix := '/read/3', Data := WORD_TO_STRING(Data^[3]));
	PubMqttMessage(Suffix := '/read/4', Data := WORD_TO_STRING(Data^[4]));
	PubMqttMessage(Suffix := '/read/5', Data := WORD_TO_STRING(Data^[5]));
END_IF
                
END_METHOD

METHOD RequestBusTime : BOOL
                  IF NOT NodeInitialized THEN	
	RequestBusTime := FALSE;
ELSIF timerData.Q THEN
	RequestBusTime := TRUE;
ELSE
	RequestBusTime := FALSE;	
END_IF
                
END_METHOD

METHOD InitNode
  VAR_INPUT
    DeviceAddress : BYTE;
    NodeNumber : UINT;
    DataPollingInterval : TIME;
  END_VAR
                  THIS^.RtuQueryRead.DeviceId := DeviceAddress;
THIS^.RtuQueryRead.ReadAddress := (NodeNumber * 10) + 10;

THIS^.timerData.PT := DataPollingInterval;
THIS^.NodeNumber := NodeNumber + 1;

THIS^.timerData.IN := TRUE;

THIS^.NodeInitialized := TRUE;
                
END_METHOD

METHOD InitMqtt
  VAR_INPUT
    MQTTPublishPrefix : POINTER TO STRING;
    MqttPublishTopicSuffix : STRING(255);
    pMqttPublishQueue : POINTER TO FB_MqttPublishQueue;
  END_VAR
                  THIS^.MqttPublishTopicPrefix := MQTTPublishPrefix;
THIS^.MqttPublishTopicSuffix := MqttPublishTopicSuffix;
THIS^.pMqttPublishQueue := pMqttPublishQueue;

THIS^.InitMqttDone := TRUE;
                
END_METHOD

METHOD PubMqttMessage
  VAR_INPUT
    Suffix : STRING(100);
    Data : STRING(100);
  END_VAR
                  IF InitMqttDone THEN
		pMqttPublishQueue^.AddMessage(
			Payload := Data,
			Topic := CONCAT(CONCAT(CONCAT(CONCAT(MqttPublishTopicPrefix^, MqttPublishTopicSuffix), '/'), UINT_TO_STRING(NodeNumber)), Suffix ),
			Qos := MQTT.QoS.ExactlyOnce,
			MqttRetain := FALSE
		);
END_IF
                
END_METHOD
END_FUNCTION_BLOCK

{attribute 'reflection'}
FUNCTION_BLOCK FB_RS485_EASTRON_SDM_POWER_MQTT IMPLEMENTS RS485Device
  VAR_OUTPUT
    ACTIVEPOWER : REAL := 0;
    DataAvailable : BOOL := FALSE;
    Error : BOOL := FALSE;
  END_VAR
  VAR
    {attribute 'instance-path'}
    {attribute 'noinit'}
    InstanceName : STRING;  (* object's full instance name *)
    Startup : BOOL := TRUE;
    InitMqttDone : BOOL;
    MqttPublishTopicPrefix : POINTER TO STRING;
    MqttPublishTopicSuffix : STRING(50);
    pMqttPublishQueue : POINTER TO FB_MqttPublishQueue;
    InitRS485Done : BOOL := FALSE;
    ActiveDevice : BOOL := FALSE;
    timerData : TON;
    isDataUpdated : BOOL := FALSE;
    DeviceType : RS485_EASTRON_SDM_Devices;
    SDM120AndSDM220RtuQuery : RS485_RtuQuery := (FunctionCode := 4, ReadAddress := 12, ReadQuantity := 2);
    SDM630RtuQuery : RS485_RtuQuery := (FunctionCode := 4, ReadAddress := 52, ReadQuantity := 2);
  END_VAR

            timerData();

IF isDataUpdated THEN
	isDataUpdated := FALSE;
	
	IF InitMqttDone THEN
		pMqttPublishQueue^.AddMessage(
			Payload := REAL_TO_STRING(ACTIVEPOWER),
			Topic := CONCAT(CONCAT(MqttPublishTopicPrefix^, MqttPublishTopicSuffix), '/ACTP' ),
			Qos := MQTT.QoS.ExactlyOnce,
			MqttRetain := FALSE
		);
	END_IF
END_IF

          

METHOD ProcessDataArray
  VAR_INPUT
    Error : POINTER TO BOOL;
    Data : POINTER TO ARRAY[0..124] OF WORD;
  END_VAR
                  THIS^.Error := Error^;
THIS^.timerData.IN := TRUE;

IF Error^ THEN
	PubMqttMessage(Suffix := '/availability', Data := 'offline');
ELSE
	PubMqttMessage(Suffix := '/availability', Data := 'online');
END_IF

IF NOT Error^ THEN
	THIS^.ACTIVEPOWER := SwapWordsToReal(Data^[0], Data^[1]);
	THIS^.isDataUpdated := TRUE;
END_IF

ActiveDevice := FALSE;




                
END_METHOD

METHOD InitRS485
  VAR_INPUT
    DataPollingInterval : TIME;
    DeviceAddress : BYTE;
    DeviceType : RS485_EASTRON_SDM_Devices;
  END_VAR
                  THIS^.timerData.PT := DataPollingInterval;
THIS^.SDM120AndSDM220RtuQuery.DeviceId := DeviceAddress;
THIS^.SDM630RtuQuery.DeviceId := DeviceAddress;
THIS^.timerData.IN := TRUE;
THIS^.DeviceType := DeviceType;

THIS^.InitRS485Done := TRUE;
                
END_METHOD

METHOD InitMqtt
  VAR_INPUT
    MQTTPublishPrefix : POINTER TO STRING;
    pMqttPublishQueue : POINTER TO FB_MqttPublishQueue;
  END_VAR
  VAR
    InstanceNamePt : POINTER TO STRING;
  END_VAR
                  THIS^.pMqttPublishQueue := pMqttPublishQueue;
THIS^.MqttPublishTopicPrefix := MQTTPublishPrefix;

InstanceNamePt := CommonTypesAndFunctions.FindLastDot(ADR(THIS^.InstanceName)) + 1;
THIS^.MqttPublishTopicSuffix := InstanceNamePt^;

THIS^.InitMqttDone := TRUE;
                
END_METHOD

METHOD RequestBusTime : BOOL
                  IF NOT InitRS485Done THEN	
	RequestBusTime := FALSE;	
ELSIF timerData.Q THEN
	RequestBusTime := TRUE;
ELSE
	RequestBusTime := FALSE;	
END_IF
                
END_METHOD

METHOD GetRtuQuery : RS485_RtuQuery
                  IF timerData.Q THEN
	THIS^.timerData.IN := FALSE;
	IF DeviceType = RS485_EASTRON_SDM_Devices.SDM120 OR  DeviceType = RS485_EASTRON_SDM_Devices.SDM220 THEN
		GetRtuQuery := THIS^.SDM120AndSDM220RtuQuery;		
	END_IF
	IF DeviceType = RS485_EASTRON_SDM_Devices.SDM630 THEN
		GetRtuQuery := THIS^.SDM630RtuQuery;		
	END_IF
END_IF
                
END_METHOD

METHOD PubMqttMessage
  VAR_INPUT
    Suffix : STRING(100);
    Data : STRING(100);
  END_VAR
                  IF InitMqttDone THEN
		pMqttPublishQueue^.AddMessage(
			Payload := Data,
			Topic := CONCAT(CONCAT(MqttPublishTopicPrefix^, MqttPublishTopicSuffix), Suffix ),
			Qos := MQTT.QoS.ExactlyOnce,
			MqttRetain := FALSE
		);
END_IF
                
END_METHOD
END_FUNCTION_BLOCK

{attribute 'reflection'}
FUNCTION_BLOCK FB_RS485_EASTRON_SDM220_MQTT IMPLEMENTS RS485Device
  VAR_OUTPUT
    VOLTAGE : REAL := 0;
    CURRENT : REAL := 0;
    ACTIVEPOWER : REAL := 0;
    APPARENT_POWER : REAL := 0;
    REACTIVE_POWER : REAL := 0;
    POWER_FACTOR : REAL := 0;
    PHASE_ANGLE : REAL := 0;
    DataAvailable1 : BOOL := FALSE;
    Error1 : BOOL := FALSE;
    FREQUENCY : REAL := 0;
    IMPORT_ACTIVE_ENERGY : REAL := 0;
    EXPORT_ACTIVE_ENERGY : REAL := 0;
    IMPORT_REACTIVE_ENERGY : REAL := 0;
    EXPORT_REACTIVE_ENERGY : REAL := 0;
    DataAvailable2 : BOOL := FALSE;
    Error2 : BOOL := FALSE;
    TOTAL_ACTIVE_ENERGY : REAL := 0;
    TOTAL_REACTIVE_ENERGY : REAL := 0;
    DataAvailable3 : BOOL := FALSE;
    Error3 : BOOL := FALSE;
  END_VAR
  VAR
    {attribute 'instance-path'}
    {attribute 'noinit'}
    InstanceName : STRING;  (* object's full instance name *)
    Startup : BOOL := TRUE;
    InitMqttDone : BOOL;
    MqttPublishTopicPrefix : POINTER TO STRING;
    MqttPublishTopicSuffix : STRING(50);
    pMqttPublishQueue : POINTER TO FB_MqttPublishQueue;
    InitRS485Done : BOOL := FALSE;
    ActiveDevice : BOOL := FALSE;
    ActiveRtuQuery : INT := 0;
    Data1RtuQuery : RS485_RtuQuery := (FunctionCode := 4, ReadAddress := 0, ReadQuantity := 40);
    Update1 : BOOL := FALSE;
    timerData1 : TON;
    Data2RtuQuery : RS485_RtuQuery := (FunctionCode := 4, ReadAddress := 70, ReadQuantity := 10);
    Update2 : BOOL := FALSE;
    timerData2 : TON;
    Data3RtuQuery : RS485_RtuQuery := (FunctionCode := 4, ReadAddress := 342, ReadQuantity := 4);
    Update3 : BOOL := FALSE;
    timerData3 : TON;
  END_VAR

            timerData1();
timerData2();
timerData3();

IF Update1 THEN
	Update1 := FALSE;
	DataAvailable1 := TRUE;
	
	IF InitMqttDone THEN
		pMqttPublishQueue^.AddMessage(
			Payload := REAL_TO_STRING(VOLTAGE),
			Topic := CONCAT(CONCAT(MqttPublishTopicPrefix^, MqttPublishTopicSuffix), '/VOLT' ),
			Qos := MQTT.QoS.ExactlyOnce,
			MqttRetain := FALSE
		);
		pMqttPublishQueue^.AddMessage(
			Payload := REAL_TO_STRING(CURRENT),
			Topic := CONCAT(CONCAT(MqttPublishTopicPrefix^, MqttPublishTopicSuffix), '/CURR' ),
			Qos := MQTT.QoS.ExactlyOnce,
			MqttRetain := FALSE
		);	
		pMqttPublishQueue^.AddMessage(
			Payload := REAL_TO_STRING(ACTIVEPOWER),
			Topic := CONCAT(CONCAT(MqttPublishTopicPrefix^, MqttPublishTopicSuffix), '/ACTP' ),
			Qos := MQTT.QoS.ExactlyOnce,
			MqttRetain := FALSE
		);
		pMqttPublishQueue^.AddMessage(
			Payload := REAL_TO_STRING(APPARENT_POWER),
			Topic := CONCAT(CONCAT(MqttPublishTopicPrefix^, MqttPublishTopicSuffix), '/APPP' ),
			Qos := MQTT.QoS.ExactlyOnce,
			MqttRetain := FALSE
		);
		pMqttPublishQueue^.AddMessage(
			Payload := REAL_TO_STRING(REACTIVE_POWER),
			Topic := CONCAT(CONCAT(MqttPublishTopicPrefix^, MqttPublishTopicSuffix), '/REAP' ),
			Qos := MQTT.QoS.ExactlyOnce,
			MqttRetain := FALSE
		);
		pMqttPublishQueue^.AddMessage(
			Payload := REAL_TO_STRING(POWER_FACTOR),
			Topic := CONCAT(CONCAT(MqttPublishTopicPrefix^, MqttPublishTopicSuffix), '/POWF' ),
			Qos := MQTT.QoS.ExactlyOnce,
			MqttRetain := FALSE
		);
		pMqttPublishQueue^.AddMessage(
			Payload := REAL_TO_STRING(PHASE_ANGLE),
			Topic := CONCAT(CONCAT(MqttPublishTopicPrefix^, MqttPublishTopicSuffix), '/PHAA' ),
			Qos := MQTT.QoS.ExactlyOnce,
			MqttRetain := FALSE
		);
	END_IF
END_IF

IF Update2 THEN
	Update2 := FALSE;
	DataAvailable2 := TRUE;
	
	IF InitMqttDone THEN
		pMqttPublishQueue^.AddMessage(
			Payload := REAL_TO_STRING(FREQUENCY),
			Topic := CONCAT(CONCAT(MqttPublishTopicPrefix^, MqttPublishTopicSuffix), '/FREQ' ),
			Qos := MQTT.QoS.ExactlyOnce,
			MqttRetain := FALSE
		);
		pMqttPublishQueue^.AddMessage(
			Payload := REAL_TO_STRING(IMPORT_ACTIVE_ENERGY),
			Topic := CONCAT(CONCAT(MqttPublishTopicPrefix^, MqttPublishTopicSuffix), '/IMAE' ),
			Qos := MQTT.QoS.ExactlyOnce,
			MqttRetain := FALSE
		);
		pMqttPublishQueue^.AddMessage(
			Payload := REAL_TO_STRING(EXPORT_ACTIVE_ENERGY),
			Topic := CONCAT(CONCAT(MqttPublishTopicPrefix^, MqttPublishTopicSuffix), '/EXAE' ),
			Qos := MQTT.QoS.ExactlyOnce,
			MqttRetain := FALSE
		);
		pMqttPublishQueue^.AddMessage(
			Payload := REAL_TO_STRING(IMPORT_REACTIVE_ENERGY),
			Topic := CONCAT(CONCAT(MqttPublishTopicPrefix^, MqttPublishTopicSuffix), '/IMRE' ),
			Qos := MQTT.QoS.ExactlyOnce,
			MqttRetain := FALSE
		);
		pMqttPublishQueue^.AddMessage(
			Payload := REAL_TO_STRING(EXPORT_REACTIVE_ENERGY),
			Topic := CONCAT(CONCAT(MqttPublishTopicPrefix^, MqttPublishTopicSuffix), '/EXRE' ),
			Qos := MQTT.QoS.ExactlyOnce,
			MqttRetain := FALSE
		);
	END_IF
END_IF

IF Update3 THEN
	Update3 := FALSE;	
	DataAvailable3 := TRUE;
	
